// ---- OTEL/TRACING/TRACESTATE/FUNCTION_BLOCKS/TraceStateFactory.TcPOU
(*
	Creates FB_TraceState values: parses a W3C tracestate header, clones a trace state, and
	truncates one to fit a carrier by the W3C rules. Like ValueFactory, every method returns
	TRUE on success, takes pDest by reference and never overwrites a pointer that is not 0.
	No trace state is a 0 pointer, so a method can succeed and leave pDest at 0.
*)
PROGRAM TraceStateFactory
VAR CONSTANT
	MAX_ENTRIES: UDINT := 32;  // W3C: at most 32 list members
	MAX_KEY_LENGTH: UDINT := 256;  // W3C key grammar
	MAX_VALUE_LENGTH: UDINT := 256;  // W3C value grammar
	MAX_HEADER_LENGTH: UDINT := 16447;  // 32 entries of the longest key and value; bounds every scan
	CARRIER_LENGTH: UDINT := 512;  // W3C: propagate at least 512 characters
	LARGE_ENTRY_LENGTH: UDINT := 128;  // W3C: when truncating, remove entries over 128 characters first
END_VAR

(*
	Allocates a trace state from the kept entries of pSource, joined by ','. Succeeds with pDest
	left at 0 when no entry is kept. The arrays are primitive scratch data owned by the caller.
*)
METHOD _build : BOOL
VAR_IN_OUT
	pDest: POINTER TO FB_TraceState;
	starts: ARRAY[0..MAX_ENTRIES - 1] OF UDINT;
	lengths: ARRAY[0..MAX_ENTRIES - 1] OF UDINT;
	keep: ARRAY[0..MAX_ENTRIES - 1] OF BOOL;
END_VAR
VAR_INPUT
	pSource: POINTER TO BYTE;
	count: UDINT;
END_VAR
VAR_OUTPUT
	failureReason: E_TraceStateFailureReason;
END_VAR
VAR
	_i: UDINT;
	_kept: UDINT;
	_length: UDINT;
	_offset: UDINT;
	_pBuffer: POINTER TO BYTE;
	_size: UDINT;
	_pNew: POINTER TO FB_TraceState;
END_VAR
_build := FALSE;
failureReason := E_TraceStateFailureReason.NA;

// size the buffer to the kept entries and the commas between them
WHILE _i < count AND _i < MAX_ENTRIES DO
	IF keep[_i] THEN
		_length := _length + lengths[_i];
		_kept := _kept + 1;
	END_IF
	_i := _i + 1;
END_WHILE
IF _kept = 0 THEN
	// nothing left is no trace state, not an empty one
	_build := TRUE;
	RETURN;
END_IF
_length := _length + _kept - 1;

_size := _length + 1;
_pBuffer := __NEW(BYTE, _size);
IF _pBuffer = 0 THEN
	failureReason := E_TraceStateFailureReason.MEMORY_ALLOCATION_FAILURE;
	RETURN;
END_IF

_i := 0;
WHILE _i < count AND _i < MAX_ENTRIES DO
	IF keep[_i] THEN
		IF _offset > 0 THEN
			_pBuffer[_offset] := 16#2C;  // ','
			_offset := _offset + 1;
		END_IF
		MEMCPY(_pBuffer + _offset, pSource + starts[_i], lengths[_i]);
		_offset := _offset + lengths[_i];
	END_IF
	_i := _i + 1;
END_WHILE
_pBuffer[_offset] := 0;

_pNew := __NEW(FB_TraceState(pString:=_pBuffer, length:=_length, count:=_kept));
IF _pNew = 0 THEN
	__DELETE(_pBuffer);
	_pBuffer := 0;
	failureReason := E_TraceStateFailureReason.MEMORY_ALLOCATION_FAILURE;
	RETURN;
END_IF
pDest := _pNew;
_build := TRUE;
END_METHOD

(* lcalpha / DIGIT / '_' / '-' / '*' / '/' *)
METHOD _isKeyChar : BOOL
VAR_INPUT
	c: BYTE;
END_VAR
_isKeyChar := (c >= 16#61 AND c <= 16#7A)  // a-z
	OR (c >= 16#30 AND c <= 16#39)  // 0-9
	OR c = 16#5F OR c = 16#2D OR c = 16#2A OR c = 16#2F;
END_METHOD

(*
	A key is either simple-key, a lower-case letter followed by up to 255 key characters, or
	multi-tenant-key: tenant-id '@' system-id, where tenant-id is 1-241 key characters starting
	with a lower-case letter or digit, and system-id is 1-14 key characters starting with a
	lower-case letter.
*)
METHOD _isValidKey : BOOL
VAR_INPUT
	pKey: POINTER TO BYTE;
	length: UDINT;
END_VAR
VAR
	_i: UDINT;
	_at: UDINT;
	_hasAt: BOOL;
	_first: BYTE;
END_VAR
_isValidKey := FALSE;
IF length = 0 OR length > MAX_KEY_LENGTH THEN
	RETURN;
END_IF

// bounded by MAX_KEY_LENGTH
WHILE _i < length DO
	IF pKey[_i] = 16#40 THEN  // '@'
		IF _hasAt THEN
			RETURN;
		END_IF
		_hasAt := TRUE;
		_at := _i;
	ELSIF NOT TraceStateFactory._isKeyChar(c:=pKey[_i]) THEN
		RETURN;
	END_IF
	_i := _i + 1;
END_WHILE

_first := pKey[0];
IF NOT _hasAt THEN
	_isValidKey := _first >= 16#61 AND _first <= 16#7A;
ELSIF _at >= 1 AND _at <= 241 AND length - _at - 1 >= 1 AND length - _at - 1 <= 14 THEN
	_isValidKey := ((_first >= 16#61 AND _first <= 16#7A) OR (_first >= 16#30 AND _first <= 16#39))
		AND pKey[_at + 1] >= 16#61 AND pKey[_at + 1] <= 16#7A;
END_IF
END_METHOD

(*
	A value is 1-256 printable ASCII characters other than ',' and '=', and does not end in a
	space.
*)
METHOD _isValidValue : BOOL
VAR_INPUT
	pValue: POINTER TO BYTE;
	length: UDINT;
END_VAR
VAR
	_i: UDINT;
	_c: BYTE;
END_VAR
_isValidValue := FALSE;
IF length = 0 OR length > MAX_VALUE_LENGTH THEN
	RETURN;
END_IF
IF pValue[length - 1] = 16#20 THEN
	RETURN;
END_IF

// bounded by MAX_VALUE_LENGTH
WHILE _i < length DO
	_c := pValue[_i];
	IF _c < 16#20 OR _c > 16#7E OR _c = 16#2C OR _c = 16#3D THEN
		RETURN;
	END_IF
	_i := _i + 1;
END_WHILE
_isValidValue := TRUE;
END_METHOD

(*
	Allocates a copy of pSrc. The caller owns pDest.
*)
METHOD clone : BOOL
VAR_IN_OUT
	pDest: POINTER TO FB_TraceState;
END_VAR
VAR_INPUT
	pSrc: POINTER TO FB_TraceState;
END_VAR
VAR_OUTPUT
	failureReason: E_TraceStateFailureReason;
END_VAR
VAR
	_pBuffer: POINTER TO BYTE;
	_size: UDINT;
	_pNew: POINTER TO FB_TraceState;
END_VAR
clone := FALSE;
failureReason := E_TraceStateFailureReason.NA;

IF pDest <> 0 THEN
	failureReason := E_TraceStateFailureReason.DESTINATION_ALREADY_ASSIGNED;
	RETURN;
END_IF
IF pSrc = 0 OR_ELSE pSrc^.pString = 0 THEN
	failureReason := E_TraceStateFailureReason.SOURCE_POINTER_NULL;
	RETURN;
END_IF

// copy by length, terminator included; the string may be longer than T_MaxString
_size := pSrc^.length + 1;
_pBuffer := __NEW(BYTE, _size);
IF _pBuffer = 0 THEN
	failureReason := E_TraceStateFailureReason.MEMORY_ALLOCATION_FAILURE;
	RETURN;
END_IF
MEMCPY(_pBuffer, pSrc^.pString, pSrc^.length + 1);

_pNew := __NEW(FB_TraceState(pString:=_pBuffer, length:=pSrc^.length, count:=pSrc^.count));
IF _pNew = 0 THEN
	__DELETE(_pBuffer);
	_pBuffer := 0;
	failureReason := E_TraceStateFailureReason.MEMORY_ALLOCATION_FAILURE;
	RETURN;
END_IF
pDest := _pNew;
clone := TRUE;
END_METHOD

(*
	Parses a W3C tracestate header into a new trace state in canonical form. The caller owns
	pDest. An empty header, or one of only empty members, is valid and succeeds with pDest left
	at 0. A header that breaks the grammar, repeats a key or has more than MAX_ENTRIES entries
	fails, and W3C says it must then not be propagated. The header may be longer than
	T_MaxString; it is measured with LEN2.
*)
METHOD parse : BOOL
VAR_IN_OUT
	pDest: POINTER TO FB_TraceState;
END_VAR
VAR_INPUT
	pHeader: POINTER TO STRING;
END_VAR
VAR_OUTPUT
	failureReason: E_TraceStateFailureReason;
END_VAR
VAR
	_pHeader: POINTER TO BYTE;
	_length: UDINT;
	_i: UDINT;
	_j: UDINT;
	_memberStart: UDINT;
	_start: UDINT;
	_end: UDINT;
	_equals: UDINT;
	_keyLength: UDINT;
	_count: UDINT;
	_starts: ARRAY[0..MAX_ENTRIES - 1] OF UDINT;
	_lengths: ARRAY[0..MAX_ENTRIES - 1] OF UDINT;
	_keyLengths: ARRAY[0..MAX_ENTRIES - 1] OF UDINT;
	_keep: ARRAY[0..MAX_ENTRIES - 1] OF BOOL;
END_VAR
parse := FALSE;
failureReason := E_TraceStateFailureReason.NA;

IF pDest <> 0 THEN
	failureReason := E_TraceStateFailureReason.DESTINATION_ALREADY_ASSIGNED;
	RETURN;
END_IF
IF pHeader = 0 THEN
	failureReason := E_TraceStateFailureReason.HEADER_POINTER_NULL;
	RETURN;
END_IF

_pHeader := pHeader;
_length := TO_UDINT(LEN2(pHeader));
IF _length > MAX_HEADER_LENGTH THEN
	failureReason := E_TraceStateFailureReason.HEADER_TOO_LONG;
	RETURN;
END_IF

// validate every member before allocating anything; _i = _length closes the last member
FOR _i := 0 TO _length DO
	IF _i < _length AND_THEN _pHeader[_i] <> 16#2C THEN  // ','
		CONTINUE;
	END_IF
	_start := _memberStart;
	_end := _i;
	_memberStart := _i + 1;

	// strip optional whitespace; an empty member is allowed and dropped
	WHILE _start < _end AND_THEN (_pHeader[_start] = 16#20 OR _pHeader[_start] = 16#09) DO
		_start := _start + 1;
	END_WHILE
	WHILE _end > _start AND_THEN (_pHeader[_end - 1] = 16#20 OR _pHeader[_end - 1] = 16#09) DO
		_end := _end - 1;
	END_WHILE
	IF _start = _end THEN
		CONTINUE;
	END_IF

	IF _count >= MAX_ENTRIES THEN
		failureReason := E_TraceStateFailureReason.TOO_MANY_ENTRIES;
		RETURN;
	END_IF

	_equals := _start;
	WHILE _equals < _end AND_THEN _pHeader[_equals] <> 16#3D DO  // '='
		_equals := _equals + 1;
	END_WHILE
	_keyLength := _equals - _start;
	IF NOT TraceStateFactory._isValidKey(pKey:=_pHeader + _start, length:=_keyLength) THEN
		failureReason := E_TraceStateFailureReason.INVALID_KEY;
		RETURN;
	END_IF
	IF _equals = _end OR_ELSE NOT TraceStateFactory._isValidValue(pValue:=_pHeader + _equals + 1, length:=_end - _equals - 1) THEN
		failureReason := E_TraceStateFailureReason.INVALID_VALUE;
		RETURN;
	END_IF

	_j := 0;
	WHILE _j < _count DO
		IF _keyLengths[_j] = _keyLength AND_THEN MEMCMP(_pHeader + _starts[_j], _pHeader + _start, _keyLength) = 0 THEN
			failureReason := E_TraceStateFailureReason.DUPLICATE_KEY;
			RETURN;
		END_IF
		_j := _j + 1;
	END_WHILE

	_starts[_count] := _start;
	_lengths[_count] := _end - _start;
	_keyLengths[_count] := _keyLength;
	_keep[_count] := TRUE;
	_count := _count + 1;
END_FOR

parse := TraceStateFactory._build(
	pDest:=pDest,
	starts:=_starts,
	lengths:=_lengths,
	keep:=_keep,
	pSource:=_pHeader,
	count:=_count,
	failureReason=>failureReason
);
END_METHOD

(*
	Allocates a copy of pSrc that is at most maxLength characters long, for a carrier of
	limited size, following W3C: entries over LARGE_ENTRY_LENGTH characters are removed first,
	then entries are removed from the right. An entry is removed whole, never cut. Succeeds with
	pDest left at 0 when no entry fits.
*)
METHOD truncate : BOOL
VAR_IN_OUT
	pDest: POINTER TO FB_TraceState;
END_VAR
VAR_INPUT
	pSrc: POINTER TO FB_TraceState;
	maxLength: UDINT;
END_VAR
VAR_OUTPUT
	failureReason: E_TraceStateFailureReason;
END_VAR
VAR
	_pSource: POINTER TO BYTE;
	_i: UDINT;
	_start: UDINT;
	_count: UDINT;
	_kept: UDINT;
	_sum: UDINT;
	_total: UDINT;
	_starts: ARRAY[0..MAX_ENTRIES - 1] OF UDINT;
	_lengths: ARRAY[0..MAX_ENTRIES - 1] OF UDINT;
	_keep: ARRAY[0..MAX_ENTRIES - 1] OF BOOL;
END_VAR
truncate := FALSE;
failureReason := E_TraceStateFailureReason.NA;

IF pDest <> 0 THEN
	failureReason := E_TraceStateFailureReason.DESTINATION_ALREADY_ASSIGNED;
	RETURN;
END_IF
IF pSrc = 0 OR_ELSE pSrc^.pString = 0 THEN
	failureReason := E_TraceStateFailureReason.SOURCE_POINTER_NULL;
	RETURN;
END_IF

IF pSrc^.length <= maxLength THEN
	truncate := TraceStateFactory.clone(pDest:=pDest, pSrc:=pSrc, failureReason=>failureReason);
	RETURN;
END_IF

// split the canonical string: entries joined by ',', no whitespace, at most MAX_ENTRIES
_pSource := pSrc^.pString;
FOR _i := 0 TO pSrc^.length DO
	IF _i = pSrc^.length OR_ELSE _pSource[_i] = 16#2C THEN
		IF _count < MAX_ENTRIES THEN
			_starts[_count] := _start;
			_lengths[_count] := _i - _start;
			_keep[_count] := TRUE;
			_sum := _sum + _i - _start;
			_count := _count + 1;
		END_IF
		_start := _i + 1;
	END_IF
END_FOR
_kept := _count;
_total := pSrc^.length;

// first remove the large entries, from the right
_i := _count;
WHILE _i > 0 AND _total > maxLength DO
	_i := _i - 1;
	IF _lengths[_i] > LARGE_ENTRY_LENGTH THEN
		_keep[_i] := FALSE;
		_sum := _sum - _lengths[_i];
		_kept := _kept - 1;
		_total := SEL(_kept > 0, 0, _sum + _kept - 1);
	END_IF
END_WHILE

// then any entry, from the right
_i := _count;
WHILE _i > 0 AND _total > maxLength DO
	_i := _i - 1;
	IF _keep[_i] THEN
		_keep[_i] := FALSE;
		_sum := _sum - _lengths[_i];
		_kept := _kept - 1;
		_total := SEL(_kept > 0, 0, _sum + _kept - 1);
	END_IF
END_WHILE

truncate := TraceStateFactory._build(
	pDest:=pDest,
	starts:=_starts,
	lengths:=_lengths,
	keep:=_keep,
	pSource:=_pSource,
	count:=_count,
	failureReason=>failureReason
);
END_METHOD

END_PROGRAM

// ---- OTEL/TRACING/SPAN/ContextFactory.TcPOU
PROGRAM ContextFactory

(*
	Allocates a span context holding copies of the given identity. The caller owns pDest.
	The identifiers are not validated; producers are responsible for what they build,
	and a context built from all-zero identifiers is simply not valid.
	pTraceState is borrowed and copied; 0 means no trace state.
*)
METHOD buildContext : BOOL
VAR_IN_OUT
	pDest: POINTER TO FB_SpanContext;
END_VAR
VAR_INPUT
	pTraceId: POINTER TO FB_TraceId;
	pSpanId: POINTER TO FB_SpanId;
	pTraceState: POINTER TO FB_TraceState;
	traceFlags: UDINT;
END_VAR
VAR_OUTPUT
	failureReason: E_ContextFactoryFailureReason;
END_VAR
VAR
	_pTraceState: POINTER TO FB_TraceState;
	_pNew: POINTER TO FB_SpanContext;
END_VAR
buildContext := FALSE;
failureReason := E_ContextFactoryFailureReason.NA;

IF pDest <> 0 THEN
	failureReason := E_ContextFactoryFailureReason.DESTINATION_ALREADY_ASSIGNED;
	RETURN;
END_IF

IF pTraceId = 0 THEN
	failureReason := E_ContextFactoryFailureReason.TRACE_ID_POINTER_NULL;
	RETURN;
END_IF

IF pSpanId = 0 THEN
	failureReason := E_ContextFactoryFailureReason.SPAN_ID_POINTER_NULL;
	RETURN;
END_IF

// clone all owned data before allocating the context itself
IF pTraceState <> 0 THEN
	IF NOT TraceStateFactory.clone(pDest:=_pTraceState, pSrc:=pTraceState) THEN
		failureReason := E_ContextFactoryFailureReason.MEMORY_ALLOCATION_FAILURE;
		RETURN;
	END_IF
END_IF

_pNew := __NEW(FB_SpanContext(
	pTraceId:=pTraceId,
	pSpanId:=pSpanId,
	pTraceState:=_pTraceState,
	traceFlags:=traceFlags
));
IF _pNew = 0 THEN
	failureReason := E_ContextFactoryFailureReason.MEMORY_ALLOCATION_FAILURE;
	IF _pTraceState <> 0 THEN _pTraceState^.delete(pSelf:=_pTraceState); END_IF
	RETURN;
END_IF
_pTraceState := 0;  // moved into FB_SpanContext
pDest := _pNew;
buildContext := failureReason = E_ContextFactoryFailureReason.NA;
END_METHOD

(*
	Allocates a snapshot of a span's identity. The caller owns pDest, which must be 0; the span
	is borrowed and unchanged. The span is the producer, and its identifiers come from the id
	generator, which only hands out valid ones, so they are not checked again here. A span that
	has not been built has no identifiers and is refused with TRACE_ID_POINTER_NULL.
	The context is always local: a span's own flags describe its parent's remoteness, so only
	the W3C trace flags are kept, and remoteness is marked as known and not remote.
*)
METHOD fromSpan : BOOL
VAR_IN_OUT
	pDest: POINTER TO FB_SpanContext;
END_VAR
VAR_INPUT
	pSpan: POINTER TO FB_Span;
END_VAR
VAR_OUTPUT
	failureReason: E_ContextFactoryFailureReason;
END_VAR
VAR
	_traceFlags: UDINT;
END_VAR
fromSpan := FALSE;
failureReason := E_ContextFactoryFailureReason.NA;

IF pSpan = 0 THEN
	failureReason := E_ContextFactoryFailureReason.SPAN_POINTER_NULL;
	RETURN;
END_IF

_traceFlags := (pSpan^.flags AND TO_UDINT(E_SpanFlags.SPAN_FLAGS_TRACE_FLAGS_MASK))
	OR TO_UDINT(E_SpanFlags.SPAN_FLAGS_CONTEXT_HAS_IS_REMOTE_MASK);

fromSpan := ContextFactory.buildContext(
	pDest:=pDest,
	pTraceId:=pSpan^.traceId,
	pSpanId:=pSpan^.spanId,
	pTraceState:=pSpan^.traceState,
	traceFlags:=_traceFlags,
	failureReason=>failureReason
);
END_METHOD

END_PROGRAM

// ---- OTEL/COMMON/FUNCTION_BLOCKS/FB_Resource.TcPOU
{attribute 'enable_dynamic_creation'}
FUNCTION_BLOCK FB_Resource
VAR_OUTPUT
	id: UDINT;	// process-local identity, assigned automatically and never exported. Snapshots share the id of their source.
	droppedAttributesCount: UDINT;
	schemaUrl: T_MaxString;
END_VAR
VAR_OUTPUT
	attributes: FB_Attributes(maxCount := TcOtlp_GVL.DEFAULT_MAX_ATTRIBUTE_COUNT);
END_VAR

METHOD copyFrom : BOOL
VAR_IN_OUT
	src: FB_Resource;
END_VAR
VAR_OUTPUT
	failureResult: E_AttributesFailureReason;
END_VAR
failureResult := E_AttributesFailureReason.NA;
THIS^.id := src.id;
THIS^.schemaUrl := src.schemaUrl;
THIS^.droppedAttributesCount := src.droppedAttributesCount;
THIS^.attributes.free();
copyFrom := THIS^.attributes.copyFrom(src:=src.attributes, failureReason=>failureResult);
END_METHOD

METHOD FB_Exit : BOOL
VAR_INPUT
	bInCopyCode: BOOL;
END_VAR
THIS^.free();
END_METHOD

//FB_Init is always available implicitly and it is used primarily for initialization.
//The return value is not evaluated. For a specific influence, you can also declare the
//methods explicitly and provide additional code there with the standard initialization
//code. You can evaluate the return value.
METHOD FB_Init: BOOL
VAR_INPUT
    bInitRetains: BOOL; // TRUE: the retain variables are initialized (reset warm / reset cold)
    bInCopyCode: BOOL;  // TRUE: the instance will be copied to the copy code afterward (online change) 
	schemaUrl: T_MaxString;
END_VAR
THIS^.schemaUrl := schemaUrl;

// claim a process-local identity; keep the existing one during an online change copy
IF NOT bInCopyCode THEN
	THIS^.id := TcOtlp_GVL.NEXT_ID;
END_IF
END_METHOD

METHOD free
THIS^.attributes.free();
END_METHOD

END_FUNCTION_BLOCK

// ---- OTEL/COMMON/FUNCTION_BLOCKS/FB_InstrumentationScope.TcPOU
FUNCTION_BLOCK FB_InstrumentationScope
VAR_OUTPUT
	name: T_MaxString;
	version: T_MaxString;
	droppedAttributesCount: UDINT;
	schemaUrl: T_MaxString;
END_VAR
VAR_OUTPUT
	attributes: FB_Attributes(maxCount := TcOtlp_GVL.DEFAULT_MAX_ATTRIBUTE_COUNT);
END_VAR

METHOD copyFrom : BOOL
VAR_IN_OUT
	src: FB_InstrumentationScope;
END_VAR
VAR_OUTPUT
	failureResult: E_AttributesFailureReason;
END_VAR
failureResult := E_AttributesFailureReason.NA;
THIS^.name := src.name;
THIS^.version := src.version;
THIS^.droppedAttributesCount := src.droppedAttributesCount;
THIS^.schemaUrl := src.schemaUrl;
THIS^.attributes.free();
copyFrom := THIS^.attributes.copyFrom(src:=src.attributes, failureReason=>failureResult);
END_METHOD

//FB_Exit must be implemented explicitly. If there is an implementation, then the
//method is called before the controller removes the code of the function block instance
//(implicit call). The return value is not evaluated.
METHOD FB_Exit: BOOL
VAR_INPUT
    bInCopyCode: BOOL;  // TRUE: the exit method is called in order to leave the instance which will be copied afterwards (online change).  
END_VAR
THIS^.free();
END_METHOD

METHOD FB_Init: BOOL
VAR_INPUT
	bInitRetains: BOOL;
	bInCopyCode: BOOL;
	name: T_MaxString;
	version: T_MaxString;
	schemaUrl: T_MaxString;
END_VAR
THIS^.name := name;
THIS^.version := version;
THIS^.schemaUrl := schemaUrl;
END_METHOD

METHOD free
VAR_INPUT
END_VAR
THIS^.attributes.free();
END_METHOD

END_FUNCTION_BLOCK

// ---- OTEL/LOGGING/EXPORTING/FUNCTION_BLOCKS/FB_LogRecordExporter_Base.TcPOU
FUNCTION_BLOCK ABSTRACT FB_LogRecordExporter_Base
VAR
	_records: FB_LogRecordQueue(maxCount:=0);
	_exportActive: BOOL;
	_callFailureReason: E_LogRecordExporterFailureReason;
END_VAR

METHOD export: BOOL
VAR_IN_OUT
	logRecords: FB_LogRecordQueue;  // accepted records are transferred out of this queue
END_VAR
VAR_INPUT
	count: UDINT;
END_VAR
VAR_OUTPUT
	failureReason: E_LogRecordExporterFailureReason;
END_VAR
VAR
	_queueFailureReason: E_LogRecordQueueFailureReason;
END_VAR
export := FALSE;
failureReason := E_LogRecordExporterFailureReason.NA;

IF THIS^.isBusy() THEN
	failureReason := E_LogRecordExporterFailureReason.ACTIVE_EXPORT_IN_PROGRESS;
	RETURN;
END_IF

// Release a completed batch retained by an exporter before accepting the next one.
THIS^.free();
IF NOT logRecords.transferTo(
	destination:=THIS^._records,
	count:=count,
	failureReason=>_queueFailureReason
) THEN
	failureReason := E_LogRecordExporterFailureReason.QUEUE_TRANSFER_FAILURE;
	RETURN;
END_IF

THIS^._exportActive := THIS^._records.count > 0;
export := failureReason = E_LogRecordExporterFailureReason.NA;
END_METHOD

METHOD FB_Exit: BOOL
VAR_INPUT
	bInCopyCode: BOOL;
END_VAR
IF NOT bInCopyCode THEN
	THIS^.free();
END_IF
END_METHOD

METHOD free
THIS^._records.free();
THIS^._exportActive := FALSE;
END_METHOD

METHOD ABSTRACT isBusy : BOOL
END_METHOD

METHOD ABSTRACT tick : BOOL
VAR_OUTPUT
	failureReason: E_LogRecordExporterFailureReason;
END_VAR
END_METHOD

END_FUNCTION_BLOCK

// ---- OTEL/LOGGING/LOG_RECORD/FUNCTION_BLOCKS/FB_LogRecordQueue.TcPOU
(*
	FIFO queue that owns every FB_LogRecord pointer it contains. push drops the
	oldest owned records when the bound is reached. The bound is maxCount, but
	never more than TcOtlp_GVL.MAX_LOOP_COUNT: a maxCount of zero, or one above
	that limit, is held to MAX_LOOP_COUNT so that free always reaches the end.
	pop transfers ownership back to the caller. transferTo moves allocated
	nodes between queue owners without copying records.
*)
FUNCTION_BLOCK FB_LogRecordQueue
VAR
	_head: POINTER TO ST_LinkedListNode;
	_tail: POINTER TO ST_LinkedListNode;
	_cursor: POINTER TO ST_LinkedListNode;
END_VAR
VAR_OUTPUT
	count: UDINT;
	maxCount: UDINT;
	droppedCount: UDINT;
END_VAR

(* The enforced bound: maxCount, held to MAX_LOOP_COUNT when it is zero or larger. *)
METHOD _capacity : UDINT
IF THIS^.maxCount = 0 OR THIS^.maxCount > TcOtlp_GVL.MAX_LOOP_COUNT THEN
	_capacity := TcOtlp_GVL.MAX_LOOP_COUNT;
ELSE
	_capacity := THIS^.maxCount;
END_IF
END_METHOD

METHOD FB_Exit : BOOL
VAR_INPUT
	bInCopyCode: BOOL;
END_VAR
IF NOT bInCopyCode THEN
	THIS^.free();
END_IF
END_METHOD

METHOD FB_Init : BOOL
VAR_INPUT
	bInitRetains: BOOL;
	bInCopyCode: BOOL;
	maxCount: UDINT := 0;
END_VAR
THIS^.maxCount := maxCount;
END_METHOD

(*
	Releases every owned record. push holds count to MAX_LOOP_COUNT, so the loop
	always reaches the end. If it ever stops early, the unreleased nodes stay in
	the queue and free returns FALSE, so a later call can finish the job.
*)
METHOD free : BOOL
VAR
	_idx: UDINT;
	_node: POINTER TO ST_LinkedListNode;
	_record: POINTER TO FB_LogRecord;
END_VAR
FOR _idx := 0 TO TcOtlp_GVL.MAX_LOOP_COUNT DO
	IF THIS^._head = 0 THEN
		EXIT;
	END_IF

	_node := THIS^._head;
	THIS^._head := _node^.nxt;
	IF _node^.val <> 0 THEN
		_record := _node^.val;
		_node^.val := 0;
		_record^.delete(pSelf:=_record);
	END_IF
	__DELETE(_node);
	IF THIS^.count > 0 THEN
		THIS^.count := THIS^.count - 1;
	END_IF
END_FOR

THIS^._cursor := THIS^._head;
IF THIS^._head = 0 THEN
	THIS^._tail := 0;
	THIS^.count := 0;
END_IF
free := THIS^._head = 0;
END_METHOD

METHOD next : POINTER TO FB_LogRecord
next := 0;

IF THIS^._cursor <> 0 THEN
	next := THIS^._cursor^.val;
	THIS^._cursor := THIS^._cursor^.nxt;
END_IF
END_METHOD

METHOD pop : BOOL
VAR_IN_OUT
	pValue: POINTER TO FB_LogRecord;
END_VAR
VAR_OUTPUT
	failureReason: E_LogRecordQueueFailureReason;
END_VAR
VAR
	_node: POINTER TO ST_LinkedListNode;
END_VAR
pop := FALSE;
failureReason := E_LogRecordQueueFailureReason.NA;

IF pValue <> 0 THEN
	failureReason := E_LogRecordQueueFailureReason.DESTINATION_ALREADY_ASSIGNED;
	RETURN;
END_IF
IF THIS^._head = 0 THEN
	failureReason := E_LogRecordQueueFailureReason.QUEUE_EMPTY;
	RETURN;
END_IF

_node := THIS^._head;
THIS^._head := _node^.nxt;
IF THIS^._cursor = _node THEN
	THIS^._cursor := THIS^._head;
END_IF
IF THIS^._head = 0 THEN
	THIS^._tail := 0;
END_IF

pValue := _node^.val;
_node^.val := 0;
_node^.nxt := 0;
__DELETE(_node);
_node := 0;
THIS^.count := THIS^.count - 1;
pop := failureReason = E_LogRecordQueueFailureReason.NA;
END_METHOD

METHOD push : BOOL
VAR_IN_OUT
	pValue: POINTER TO FB_LogRecord;
END_VAR
VAR_OUTPUT
	failureReason: E_LogRecordQueueFailureReason;
END_VAR
VAR
	_node: POINTER TO ST_LinkedListNode;
	_droppedRecord: POINTER TO FB_LogRecord;
	_popFailureReason: E_LogRecordQueueFailureReason;
	_idx: UDINT;
	_bound: UDINT;
END_VAR
push := FALSE;
failureReason := E_LogRecordQueueFailureReason.NA;

IF pValue = 0 THEN
	failureReason := E_LogRecordQueueFailureReason.RECORD_POINTER_NULL;
	RETURN;
END_IF

// Allocate before evicting so an allocation failure leaves the queue unchanged.
_node := __NEW(ST_LinkedListNode);
IF _node = 0 THEN
	failureReason := E_LogRecordQueueFailureReason.MEMORY_ALLOCATION_FAILURE;
	RETURN;
END_IF

// maxCount is writable, so also restore the bound after a runtime reduction.
_bound := THIS^._capacity();
FOR _idx := 0 TO TcOtlp_GVL.MAX_LOOP_COUNT DO
	IF THIS^.count < _bound THEN
		EXIT;
	END_IF
	IF NOT THIS^.pop(pValue:=_droppedRecord, failureReason=>_popFailureReason) THEN
		__DELETE(_node);
		_node := 0;
		failureReason := _popFailureReason;
		RETURN;
	END_IF
	_droppedRecord^.delete(pSelf:=_droppedRecord);
	THIS^.droppedCount := THIS^.droppedCount + 1;
END_FOR
IF THIS^.count >= _bound THEN
	__DELETE(_node);
	_node := 0;
	failureReason := E_LogRecordQueueFailureReason.MAX_SIZE_ENFORCEMENT_FAILURE;
	RETURN;
END_IF

_node^.val := pValue;
_node^.nxt := 0;
IF THIS^._tail = 0 THEN
	THIS^._head := _node;
	THIS^._cursor := _node;
ELSE
	THIS^._tail^.nxt := _node;
END_IF
THIS^._tail := _node;
THIS^.count := THIS^.count + 1;
pValue := 0;
push := failureReason = E_LogRecordQueueFailureReason.NA;
END_METHOD

METHOD reset
THIS^._cursor := THIS^._head;
END_METHOD

(* Moves the head node to the tail without changing record ownership. *)
METHOD rotate : BOOL
VAR_OUTPUT
	failureReason: E_LogRecordQueueFailureReason;
END_VAR
VAR
	_node: POINTER TO ST_LinkedListNode;
END_VAR
rotate := FALSE;
failureReason := E_LogRecordQueueFailureReason.NA;

IF THIS^._head = 0 THEN
	failureReason := E_LogRecordQueueFailureReason.QUEUE_EMPTY;
	RETURN;
END_IF

IF THIS^._head <> THIS^._tail THEN
	_node := THIS^._head;
	THIS^._head := _node^.nxt;
	_node^.nxt := 0;
	THIS^._tail^.nxt := _node;
	THIS^._tail := _node;
END_IF

THIS^._cursor := THIS^._head;
rotate := failureReason = E_LogRecordQueueFailureReason.NA;
END_METHOD

(*
	Transfers the allocated nodes and owned records without copying them.
	The destination must be a different, empty queue. It receives up to count
	of the oldest records, also respecting the destination's bound.
*)
METHOD transferTo : BOOL
VAR_IN_OUT
	destination: FB_LogRecordQueue;
END_VAR
VAR_INPUT
	count: UDINT;
END_VAR
VAR_OUTPUT
	failureReason: E_LogRecordQueueFailureReason;
END_VAR
VAR
	_transferCount: UDINT;
	_idx: UDINT;
END_VAR
transferTo := FALSE;
failureReason := E_LogRecordQueueFailureReason.NA;

IF ADR(destination) = THIS THEN
	failureReason := E_LogRecordQueueFailureReason.SELF_TRANSFER_NOT_ALLOWED;
	RETURN;
END_IF
IF destination.count <> 0 OR_ELSE destination._head <> 0 OR_ELSE destination._tail <> 0 THEN
	failureReason := E_LogRecordQueueFailureReason.DESTINATION_NOT_EMPTY;
	RETURN;
END_IF

_transferCount := count;
IF _transferCount > THIS^.count THEN
	_transferCount := THIS^.count;
END_IF
IF _transferCount > destination._capacity() THEN
	_transferCount := destination._capacity();
END_IF
IF _transferCount = 0 THEN
	transferTo := failureReason = E_LogRecordQueueFailureReason.NA;
	RETURN;
END_IF

destination._head := THIS^._head;
destination._tail := destination._head;
FOR _idx := 1 TO _transferCount - 1 DO
	destination._tail := destination._tail^.nxt;
END_FOR

THIS^._head := destination._tail^.nxt;
destination._tail^.nxt := 0;
destination._cursor := destination._head;
destination.count := _transferCount;

THIS^.count := THIS^.count - _transferCount;
THIS^._cursor := THIS^._head;
IF THIS^._head = 0 THEN
	THIS^._tail := 0;
END_IF
transferTo := failureReason = E_LogRecordQueueFailureReason.NA;
END_METHOD

END_FUNCTION_BLOCK

// ---- OTEL/LOGGING/LOG_RECORD/FUNCTION_BLOCKS/FB_LogRecord.TcPOU
{attribute 'enable_dynamic_creation'}
FUNCTION_BLOCK FB_LogRecord
VAR_INPUT
	// required values
	severityNumber: E_SeverityNumber;
	timestamp: 		ULINT;
	
	// optional values
	eventName: 	POINTER TO FB_String; 
	traceId: 	POINTER TO FB_TraceId;
	spanId: 	POINTER TO FB_SpanId;
	flags: UDINT;  // OTLP fixed32: bits 0-7 are the W3C trace flags of the record's span (bit 0 is sampled), bits 8-31 are reserved
	body: 		POINTER TO FB_AnyValue;
	droppedAttributesCount: UDINT;
END_VAR
VAR_OUTPUT
	resource: FB_Resource('');
	scope: FB_InstrumentationScope('', '', '');
	attributes: FB_Attributes(maxCount := TcOtlp_GVL.DEFAULT_MAX_ATTRIBUTE_COUNT);
END_VAR

METHOD cloneTo : BOOL
VAR_IN_OUT
	pDest: POINTER TO FB_LogRecord;
END_VAR
VAR_OUTPUT
	failureReason: E_LogRecordCloneFailureReason;
END_VAR
VAR
	_pClone: POINTER TO FB_LogRecord;
	_factoryFailureReason: E_ValueFactoryFailureReason;
	_attributesFailureReason: E_AttributesFailureReason;
END_VAR
cloneTo := FALSE;
failureReason := E_LogRecordCloneFailureReason.NA;

IF pDest <> 0 THEN
	failureReason := E_LogRecordCloneFailureReason.DESTINATION_ALREADY_ASSIGNED;
	RETURN;
END_IF

_pClone := __NEW(FB_LogRecord(
	severityNumber:=THIS^.severityNumber,
	timestamp:=THIS^.timestamp
));
IF _pClone = 0 THEN
	failureReason := E_LogRecordCloneFailureReason.MEMORY_ALLOCATION_FAILURE;
	RETURN;
END_IF

_pClone^.droppedAttributesCount := THIS^.droppedAttributesCount;
_pClone^.flags := THIS^.flags;

IF THIS^.eventName <> 0 THEN
	IF NOT ValueFactory.cloneString(
		pDest:=_pClone^.eventName,
		pSrc:=THIS^.eventName,
		failureReason=>_factoryFailureReason
	) THEN
		IF _factoryFailureReason = E_ValueFactoryFailureReason.MEMORY_ALLOCATION_FAILURE THEN
			failureReason := E_LogRecordCloneFailureReason.MEMORY_ALLOCATION_FAILURE;
		ELSE
			failureReason := E_LogRecordCloneFailureReason.EVENT_NAME_INVALID;
		END_IF
		_pClone^.delete(pSelf:=_pClone);
		RETURN;
	END_IF
END_IF

IF THIS^.traceId <> 0 THEN
	IF NOT ValueFactory.createTraceId(
		pDest:=_pClone^.traceId,
		pBytes:=ADR(THIS^.traceId^.bytes),
		nSize:=SIZEOF(THIS^.traceId^.bytes),
		failureReason=>_factoryFailureReason
	) THEN
		IF _factoryFailureReason = E_ValueFactoryFailureReason.MEMORY_ALLOCATION_FAILURE THEN
			failureReason := E_LogRecordCloneFailureReason.MEMORY_ALLOCATION_FAILURE;
		ELSE
			failureReason := E_LogRecordCloneFailureReason.TRACE_ID_INVALID;
		END_IF
		_pClone^.delete(pSelf:=_pClone);
		RETURN;
	END_IF
END_IF

IF THIS^.spanId <> 0 THEN
	IF NOT ValueFactory.createSpanId(
		pDest:=_pClone^.spanId,
		pBytes:=ADR(THIS^.spanId^.bytes),
		nSize:=SIZEOF(THIS^.spanId^.bytes),
		failureReason=>_factoryFailureReason
	) THEN
		IF _factoryFailureReason = E_ValueFactoryFailureReason.MEMORY_ALLOCATION_FAILURE THEN
			failureReason := E_LogRecordCloneFailureReason.MEMORY_ALLOCATION_FAILURE;
		ELSE
			failureReason := E_LogRecordCloneFailureReason.SPAN_ID_INVALID;
		END_IF
		_pClone^.delete(pSelf:=_pClone);
		RETURN;
	END_IF
END_IF

IF THIS^.body <> 0 THEN
	IF NOT ValueFactory.cloneAnyValue(
		pDest:=_pClone^.body,
		pSrc:=THIS^.body,
		failureReason=>_factoryFailureReason
	) THEN
		CASE _factoryFailureReason OF
			E_ValueFactoryFailureReason.MEMORY_ALLOCATION_FAILURE:
				failureReason := E_LogRecordCloneFailureReason.MEMORY_ALLOCATION_FAILURE;
			E_ValueFactoryFailureReason.UNSUPPORTED_VALUE_TYPE:
				failureReason := E_LogRecordCloneFailureReason.BODY_VALUE_TYPE_UNSUPPORTED;
		ELSE
			failureReason := E_LogRecordCloneFailureReason.BODY_VALUE_INVALID;
		END_CASE
		_pClone^.delete(pSelf:=_pClone);
		RETURN;
	END_IF
END_IF

IF NOT _pClone^.resource.copyFrom(src:=THIS^.resource, failureResult=>_attributesFailureReason) THEN
	IF _attributesFailureReason = E_AttributesFailureReason.MEMORY_ALLOCATION_FAILURE THEN
		failureReason := E_LogRecordCloneFailureReason.MEMORY_ALLOCATION_FAILURE;
	ELSE
		failureReason := E_LogRecordCloneFailureReason.RESOURCE_COPY_FAILURE;
	END_IF
	_pClone^.delete(pSelf:=_pClone);
	RETURN;
END_IF

IF NOT _pClone^.scope.copyFrom(src:=THIS^.scope, failureResult=>_attributesFailureReason) THEN
	IF _attributesFailureReason = E_AttributesFailureReason.MEMORY_ALLOCATION_FAILURE THEN
		failureReason := E_LogRecordCloneFailureReason.MEMORY_ALLOCATION_FAILURE;
	ELSE
		failureReason := E_LogRecordCloneFailureReason.SCOPE_COPY_FAILURE;
	END_IF
	_pClone^.delete(pSelf:=_pClone);
	RETURN;
END_IF

IF NOT _pClone^.attributes.copyFrom(
	src:=THIS^.attributes,
	failureReason=>_attributesFailureReason
	) THEN
	IF _attributesFailureReason = E_AttributesFailureReason.MEMORY_ALLOCATION_FAILURE THEN
		failureReason := E_LogRecordCloneFailureReason.MEMORY_ALLOCATION_FAILURE;
	ELSE
		failureReason := E_LogRecordCloneFailureReason.ATTRIBUTE_COPY_FAILURE;
	END_IF
	_pClone^.delete(pSelf:=_pClone);
	RETURN;
END_IF

pDest := _pClone;
_pClone := 0;
cloneTo := failureReason = E_LogRecordCloneFailureReason.NA;
END_METHOD

(*
	Releases this record and clears the caller's pointer to it: call it as p^.delete(pSelf:=p).
	pSelf is cleared before the record is freed, so the caller never keeps a dangling pointer.
	A pointer to any other object is refused and left untouched, and nothing is released.
*)
METHOD delete : BOOL
VAR_IN_OUT
	pSelf: POINTER TO FB_LogRecord;
END_VAR
VAR
	_pThis: POINTER TO FB_LogRecord;
END_VAR
_pThis := THIS;
IF pSelf <> _pThis THEN
	RETURN;
END_IF

pSelf := 0;
__DELETE(_pThis);
delete := TRUE;
END_METHOD

//FB_Exit must be implemented explicitly. If there is an implementation, then the
//method is called before the controller removes the code of the function block instance
//(implicit call). The return value is not evaluated.
METHOD FB_Exit: BOOL
VAR_INPUT
    bInCopyCode: BOOL;  // TRUE: the exit method is called in order to leave the instance which will be copied afterwards (online change).
END_VAR
IF NOT bInCopyCode THEN
	THIS^.free();
END_IF
END_METHOD

//FB_Init is always available implicitly and it is used primarily for initialization.
//The return value is not evaluated. For a specific influence, you can also declare the
//methods explicitly and provide additional code there with the standard initialization
//code. You can evaluate the return value.
METHOD FB_Init: BOOL
VAR_INPUT
    bInitRetains: BOOL; // TRUE: the retain variables are initialized (reset warm / reset cold)
    bInCopyCode: BOOL;  // TRUE: the instance will be copied to the copy code afterward (online change)
	// required values
	severityNumber: E_SeverityNumber;
	timestamp: 		ULINT;
END_VAR
// required values
THIS^.severityNumber := severityNumber;
THIS^.timestamp := timestamp;
END_METHOD

METHOD free
IF THIS^.eventName <> 0 THEN THIS^.eventName^.delete(pSelf:=THIS^.eventName); END_IF
IF THIS^.traceId <> 0 THEN THIS^.traceId^.delete(pSelf:=THIS^.traceId); END_IF
IF THIS^.spanId <> 0 THEN THIS^.spanId^.delete(pSelf:=THIS^.spanId); END_IF
IF THIS^.body <> 0 THEN THIS^.body^.delete(pSelf:=THIS^.body); END_IF
THIS^.attributes.free();
THIS^.scope.free();
THIS^.resource.free();
END_METHOD

PROPERTY severityText : STRING(30)
GET
severityText := TO_STRING(THIS^.severityNumber);
END_GET
END_PROPERTY

END_FUNCTION_BLOCK

// ---- OTEL/LOGGING/EXPORTING/FUNCTION_BLOCKS/FB_LogRecordExporter_Console.TcPOU
FUNCTION_BLOCK FB_LogRecordExporter_Console EXTENDS FB_LogRecordExporter_Base
VAR_INPUT
END_VAR
VAR_OUTPUT
END_VAR
VAR
END_VAR

THIS^.tick(failureReason=>THIS^._callFailureReason);

METHOD export : BOOL
VAR_IN_OUT
	logRecords: FB_LogRecordQueue;
END_VAR
VAR_INPUT
	count: UDINT;
END_VAR
VAR_OUTPUT
	failureReason: E_LogRecordExporterFailureReason;
END_VAR
export := SUPER^.export(
	logRecords:=logRecords,
	count:=count,
	failureReason=>failureReason
);
IF NOT export THEN
	RETURN;
END_IF

THIS^.writeToConsole(THIS^._records);
THIS^.free();
END_METHOD

METHOD isBusy : BOOL
isBusy := FALSE;
END_METHOD

METHOD tick : BOOL
VAR_OUTPUT
	failureReason: E_LogRecordExporterFailureReason;
END_VAR
failureReason := E_LogRecordExporterFailureReason.NA;
tick := TRUE;
END_METHOD

METHOD writeToConsole
VAR_IN_OUT
	logRecords: FB_LogRecordQueue;
END_VAR
VAR
	idx: DINT;
	logRecord: POINTER TO FB_LogRecord;
	body: POINTER TO FB_String;
END_VAR
logRecords.reset();
FOR idx := 0 TO TcOtlp_GVL.MAX_LOOP_COUNT DO
	logRecord := logRecords.next();
	IF logRecord = 0 THEN
		RETURN;
	END_IF
	IF logRecord^.body <> 0 AND_THEN logRecord^.body^.eType = E_ValueType.E_String THEN
		body := logRecord^.body;
		ADSLOGSTR(
			ADSLOG_MSGTYPE_ERROR,
			body^.pString^,
			''
		);
	END_IF
END_FOR
END_METHOD

END_FUNCTION_BLOCK

// ---- OTEL/LOGGING/EXPORTING/FUNCTION_BLOCKS/FB_LogRecordExporter_File.TcPOU
FUNCTION_BLOCK FB_LogRecordExporter_File EXTENDS FB_LogRecordExporter_Base
VAR_INPUT
	// maxFileSize: 	UDINT;  // size at which to auto rotate the file
	// maxFiles: 		UDINT;  // max number of files to keep in the rotation
END_VAR

VAR_OUTPUT
	currentState: E_FileExporterState;
END_VAR

VAR
	_execute: BOOL;
	_filepath: T_MaxString;
	_hFile: UINT;
	_len: UDINT;
	_execRTrig: R_TRIG;
	_pString: POINTER TO STRING;
	_jsonVal: SJsonValue;
	_resourceLogsArray: SJsonValue;
	_fileOpener: FB_FileOpen;
	_fileWriter: FB_FileWrite;
	_fileCloser: FB_FileClose;
	_computedState: E_FileExporterState;
	_failureReason: E_LogRecordExporterFailureReason;
	_serializationFailureReason: E_ProtoJsonSerializerFailureReason;
	_serializer: FB_LogRecordProtoJsonSerializer;
END_VAR

THIS^.tick(failureReason=>THIS^._callFailureReason);

METHOD export: BOOL
VAR_IN_OUT
	logRecords: FB_LogRecordQueue;
END_VAR
VAR_INPUT
	count: UDINT;
END_VAR
VAR_OUTPUT
	failureReason: E_LogRecordExporterFailureReason;
END_VAR
// Prepare a completed exporter to accept the next batch immediately.
IF THIS^.currentState = E_FileExporterState.done OR THIS^.currentState = E_FileExporterState.error THEN
	THIS^.currentState := E_FileExporterState.idle;
	THIS^._computedState := E_FileExporterState.idle;
END_IF
export := SUPER^.export(
	logRecords:=logRecords,
	count:=count,
	failureReason=>failureReason
);
IF export THEN
	THIS^._failureReason := E_LogRecordExporterFailureReason.NA;
	THIS^._serializationFailureReason := E_ProtoJsonSerializerFailureReason.NA;
END_IF
END_METHOD

(*
	Releases a payload buffer that is still in flight. The FB_FileWrite reading it is
	destroyed with this instance, so nothing uses the buffer afterwards. TwinCAT then
	runs FB_LogRecordExporter_Base.FB_Exit, which releases the queued records.
*)
METHOD FB_Exit : BOOL
VAR_INPUT
	bInCopyCode: BOOL;  // TRUE: the instance is being copied during an online change
END_VAR
// during an online change the copy keeps the buffer, so it must not be released here
IF NOT bInCopyCode AND _pString <> 0 THEN
	__DELETE(_pString);
	_pString := 0;
END_IF
END_METHOD

//FB_Init is always available implicitly and it is used primarily for initialization.
//The return value is not evaluated. For a specific influence, you can also declare the
//methods explicitly and provide additional code there with the standard initialization
//code. You can evaluate the return value.
METHOD FB_Init: BOOL
VAR_INPUT
    bInitRetains: BOOL; // TRUE: the retain variables are initialized (reset warm / reset cold)
    bInCopyCode: BOOL;  // TRUE: the instance will be copied to the copy code afterward (online change)
	filepath: T_MaxString;  // path to the root file
END_VAR
THIS^._filepath := filepath;
END_METHOD

METHOD isBusy : BOOL
isBusy := THIS^._exportActive;
END_METHOD

METHOD tick : BOOL
VAR_OUTPUT
	failureReason: E_LogRecordExporterFailureReason;
END_VAR
tick := TRUE;
failureReason := E_LogRecordExporterFailureReason.NA;

_execute := THIS^._exportActive;
_execRTrig(CLK := _execute AND_THEN THIS^._records.count > 0);

CASE currentState OF
	E_FileExporterState.idle:
		IF _execRTrig.Q THEN
			_failureReason := E_LogRecordExporterFailureReason.NA;
			_serializationFailureReason := E_ProtoJsonSerializerFailureReason.NA;
			_computedState := E_FileExporterState.serializing;
		END_IF

	E_FileExporterState.serializing:
		IF NOT _serializer.serializeLogsData(
			logRecords:=THIS^._records,
			failureReason=>_serializationFailureReason
		) THEN
			_failureReason := E_LogRecordExporterFailureReason.SERIALIZATION_FAILURE;
			_computedState := E_FileExporterState.error;
		ELSE
			_jsonVal := _serializer.jsonValue;
			IF _jsonVal = 0 OR_ELSE NOT _serializer.parser.IsObject(_jsonVal) THEN
				_failureReason := E_LogRecordExporterFailureReason.SERIALIZATION_FAILURE;
				_computedState := E_FileExporterState.error;
			ELSE
				_resourceLogsArray := _serializer.parser.FindMember(_jsonVal, 'resourceLogs');
				IF _resourceLogsArray = 0 OR_ELSE NOT _serializer.parser.IsArray(_resourceLogsArray) THEN
					_failureReason := E_LogRecordExporterFailureReason.SERIALIZATION_FAILURE;
					_computedState := E_FileExporterState.error;
				ELSE
					_computedState := E_FileExporterState.opening;
				END_IF
			END_IF
		END_IF

	E_FileExporterState.opening:
		IF _fileOpener.bError THEN
			_failureReason := E_LogRecordExporterFailureReason.FILE_OPEN_FAILURE;
			_computedState := E_FileExporterState.error;
		ELSIF NOT _fileOpener.bBusy THEN
			_hFile := _fileOpener.hFile;
			_computedState := E_FileExporterState.buffering;
		END_IF

	E_FileExporterState.buffering:
		// Write one complete LogsData object per JSONL line.
		_len := _serializer.parser.GetJsonLength(_jsonVal);  // includes the null terminating character
		IF _len = 0 THEN
			_failureReason := E_LogRecordExporterFailureReason.SERIALIZATION_FAILURE;
			_computedState := E_FileExporterState.closing;
		ELSE
			_pString := __NEW(BYTE, (_len + 1));  // + 1 for the new line
			IF _pString = 0 THEN
				_failureReason := E_LogRecordExporterFailureReason.BUFFER_ALLOCATION_FAILURE;
				_computedState := E_FileExporterState.closing;
			ELSE
				_serializer.parser.CopyJson(_jsonVal, _pString^, _len);
				CONCAT2(_pString, ADR('$N'), _pString, _len + 1);
				_computedState := E_FileExporterState.writing;
			END_IF
		END_IF

	E_FileExporterState.writing:
		IF _fileWriter.bError THEN
			IF _pString <> 0 THEN __DELETE(_pString); _pString := 0; END_IF
			_failureReason := E_LogRecordExporterFailureReason.FILE_WRITE_FAILURE;
			_computedState := E_FileExporterState.closing;
		ELSIF NOT _fileWriter.bBusy THEN
			IF _pString <> 0 THEN __DELETE(_pString); _pString := 0; END_IF
			_computedState := E_FileExporterState.closing;
		END_IF

	E_FileExporterState.closing:
		IF _fileCloser.bError THEN
			IF _failureReason = E_LogRecordExporterFailureReason.NA THEN
				_failureReason := E_LogRecordExporterFailureReason.FILE_CLOSE_FAILURE;
			END_IF
			_computedState := E_FileExporterState.error;
		ELSIF NOT _fileCloser.bBusy THEN
			IF _failureReason = E_LogRecordExporterFailureReason.NA THEN
				_computedState := E_FileExporterState.done;
			ELSE
				_computedState := E_FileExporterState.error;
			END_IF
		END_IF

	E_FileExporterState.done:
		IF NOT _execute THEN
			_computedState := E_FileExporterState.idle;
		END_IF
		THIS^.free();

	E_FileExporterState.error:
		// Retain the failure until export accepts a new batch.
END_CASE

currentState := _computedState;

IF currentState <= E_FileExporterState.serializing THEN _hFile := 0; END_IF
IF currentState = E_FileExporterState.done
	OR_ELSE currentState = E_FileExporterState.error THEN
	THIS^.free();
END_IF

_fileOpener(
	sNetId:='',
	sPathName:=THIS^._filepath,
	bExecute:=currentState = E_FileExporterState.opening,
	nMode:=FOPEN_MODEAPPEND OR FOPEN_MODETEXT,
	ePath:=PATH_GENERIC,
	tTimeout:=DEFAULT_ADS_TIMEOUT
);

_fileWriter(
	hFile:=_hFile,
	bExecute:=currentState = E_FileExporterState.writing,
	pWriteBuff:=_pString,
	cbWriteLen:=_len
);

_fileCloser(
	hFile:=_hFile,
	bExecute:=currentState = E_FileExporterState.closing
);

IF currentState = E_FileExporterState.error THEN
	tick := FALSE;
	failureReason := _failureReason;
END_IF
END_METHOD

END_FUNCTION_BLOCK

// ---- OTEL/LOGGING/SERIALIZATION/FUNCTION_BLOCKS/FB_LogRecordProtoJsonSerializer.TcPOU
FUNCTION_BLOCK FB_LogRecordProtoJsonSerializer EXTENDS FB_BaseProtoJsonSerializer

METHOD serializeLogRecord : BOOL
VAR_IN_OUT
	v: SJsonValue;
END_VAR
VAR_INPUT
	pLogRecord: POINTER TO FB_LogRecord;
END_VAR
VAR_OUTPUT
	failureReason: E_ProtoJsonSerializerFailureReason;
END_VAR
VAR
	_buf: T_MaxString;
	_obj: SJsonValue;
	_member: SJsonValue;
END_VAR
serializeLogRecord := FALSE;
failureReason := E_ProtoJsonSerializerFailureReason.NA;
IF v = 0 THEN
	failureReason := E_ProtoJsonSerializerFailureReason.JSON_VALUE_INVALID;
	RETURN;
END_IF
IF pLogRecord = 0 THEN
	failureReason := E_ProtoJsonSerializerFailureReason.LOG_RECORD_POINTER_NULL;
	RETURN;
END_IF

_obj := THIS^.parser.PushbackJsonValue(v, '{}');
IF _obj = 0 THEN
	failureReason := E_ProtoJsonSerializerFailureReason.JSON_OPERATION_FAILURE;
	RETURN;
END_IF

_buf := pLogRecord^.severityText;
_member := THIS^.parser.AddUintMember(_obj, 'severityNumber', TO_UDINT(pLogRecord^.severityNumber));
IF _member = 0 THEN failureReason := E_ProtoJsonSerializerFailureReason.JSON_OPERATION_FAILURE; RETURN; END_IF
_member := THIS^.parser.AddStringMember(_obj, 'severityText', _buf);
IF _member = 0 THEN failureReason := E_ProtoJsonSerializerFailureReason.JSON_OPERATION_FAILURE; RETURN; END_IF
IF NOT THIS^.serializeUint64Value(_obj, ADR('timeUnixNano'), pLogRecord^.timestamp, failureReason=>failureReason) THEN RETURN; END_IF

IF pLogRecord^.eventName <> 0 AND_THEN NOT THIS^.serializeStringValue(_obj, ADR('eventName'), pLogRecord^.eventName, failureReason=>failureReason) THEN RETURN; END_IF
IF pLogRecord^.traceId <> 0 AND_THEN NOT THIS^.serializeTraceIdValue(_obj, pLogRecord^.traceId, failureReason=>failureReason) THEN RETURN; END_IF
IF pLogRecord^.traceId <> 0 AND_THEN NOT THIS^.serializeUint32Value(_obj, ADR('flags'), TO_UDINT(pLogRecord^.flags), failureReason=>failureReason) THEN RETURN; END_IF
IF pLogRecord^.spanId <> 0 AND_THEN NOT THIS^.serializeSpanIdValue(_obj, pLogRecord^.spanId, failureReason=>failureReason) THEN RETURN; END_IF
IF pLogRecord^.body <> 0 AND_THEN NOT THIS^.serializeAnyValue(_obj, ADR('body'), pLogRecord^.body, failureReason=>failureReason) THEN RETURN; END_IF
IF pLogRecord^.attributes.count > 0 AND_THEN NOT THIS^.serializeKeyValues(_obj, ADR('attributes'), ADR(pLogRecord^.attributes), failureReason=>failureReason) THEN RETURN; END_IF
IF pLogRecord^.droppedAttributesCount > 0 AND_THEN NOT THIS^.serializeUint32Value(
	_obj,
	ADR('droppedAttributesCount'),
	pLogRecord^.droppedAttributesCount,
	failureReason=>failureReason
) THEN
	RETURN;
END_IF
serializeLogRecord := failureReason = E_ProtoJsonSerializerFailureReason.NA;
END_METHOD

(*
	Takes ownership of all supplied records. Popped records and records remaining in the
	queue are released on both success and failure.
*)
METHOD serializeLogsData : BOOL
VAR_IN_OUT
	logRecords: FB_LogRecordQueue;
END_VAR
VAR_OUTPUT
	failureReason: E_ProtoJsonSerializerFailureReason;
END_VAR
VAR
	_ownedRecordCount: UDINT;
	_pOwnedRecord: POINTER TO FB_LogRecord;
	_resourceLogs: SJsonValue;
	_resourceIdx: UDINT;
	_queueFailureReason: E_LogRecordQueueFailureReason;
END_VAR
serializeLogsData := FALSE;
failureReason := E_ProtoJsonSerializerFailureReason.NA;

// fail early if loop limit exceeded.
_ownedRecordCount := logRecords.count;
IF _ownedRecordCount > TcOtlp_GVL.MAX_LOOP_COUNT THEN
	logRecords.free();
	failureReason := E_ProtoJsonSerializerFailureReason.LOOP_LIMIT_EXCEEDED;
	RETURN;
END_IF

// start a new document in make the first entry an object i.e. "{}"
THIS^.jsonValue := THIS^.parser.NewDocument();
IF THIS^.jsonValue = 0 THEN
	logRecords.free();
	failureReason := E_ProtoJsonSerializerFailureReason.JSON_OPERATION_FAILURE;
	RETURN;
END_IF
THIS^.jsonValue := THIS^.parser.SetObject(THIS^.jsonValue);
IF THIS^.jsonValue = 0 THEN
	logRecords.free();
	failureReason := E_ProtoJsonSerializerFailureReason.JSON_OPERATION_FAILURE;
	RETURN;
END_IF

// start the resource logs block
_resourceLogs := THIS^.parser.AddArrayMember(THIS^.jsonValue, 'resourceLogs', 0);
IF _resourceLogs = 0 THEN
	logRecords.free();
	failureReason := E_ProtoJsonSerializerFailureReason.JSON_OPERATION_FAILURE;
	RETURN;
END_IF

_pOwnedRecord := 0;
IF _ownedRecordCount > 0 THEN
	FOR _resourceIdx := 1 TO _ownedRecordCount DO
		IF logRecords.count = 0 THEN EXIT; END_IF

		// pop the record to start the group
		IF NOT logRecords.pop(pValue:=_pOwnedRecord, failureReason=>_queueFailureReason) THEN
			failureReason := E_ProtoJsonSerializerFailureReason.QUEUE_POP_FAILURE;
			EXIT;
		END_IF
		IF _pOwnedRecord = 0 THEN
			failureReason := E_ProtoJsonSerializerFailureReason.LOG_RECORD_COLLECTION_INCONSISTENT;
			EXIT;
		END_IF

		// Recursively descend from LogsData into ResourceLogs and ScopeLogs.
		IF NOT THIS^.serializeResourceLogs(
			v:=_resourceLogs,
			logRecords:=logRecords,
			pLogRecord:=_pOwnedRecord,
			failureReason=>failureReason
		) THEN
			EXIT;
		END_IF
	END_FOR
END_IF

// clean up the last record if it's not cleaned up already
IF _pOwnedRecord <> 0 THEN
	_pOwnedRecord^.delete(pSelf:=_pOwnedRecord);
END_IF

// set flag if log records didn't all get consumed
IF logRecords.count > 0 THEN
	failureReason := E_ProtoJsonSerializerFailureReason.LOOP_LIMIT_EXCEEDED;
END_IF

// free all the memory and return status
logRecords.free();
serializeLogsData := failureReason = E_ProtoJsonSerializerFailureReason.NA;
END_METHOD

METHOD serializeResourceLogs : BOOL
VAR_IN_OUT
	v: SJsonValue;
	logRecords: FB_LogRecordQueue;
	pLogRecord: POINTER TO FB_LogRecord;
END_VAR
VAR_OUTPUT
	failureReason: E_ProtoJsonSerializerFailureReason;
END_VAR
VAR
	_resourceId: UDINT;
	_scopeLogs: SJsonValue;
	_pHeadRecord: POINTER TO FB_LogRecord;
	_scopeLimit: UDINT;
	_recordsToScan: UDINT;
	_scopeIdx: UDINT;
	_scanIdx: UDINT;
	_queueFailureReason: E_LogRecordQueueFailureReason;
END_VAR
serializeResourceLogs := FALSE;
failureReason := E_ProtoJsonSerializerFailureReason.NA;
IF v = 0 THEN
	failureReason := E_ProtoJsonSerializerFailureReason.JSON_VALUE_INVALID;
	RETURN;
END_IF
IF pLogRecord = 0 THEN
	failureReason := E_ProtoJsonSerializerFailureReason.LOG_RECORD_POINTER_NULL;
	RETURN;
END_IF

_resourceId := pLogRecord^.resource.id;
IF NOT THIS^.startNewResource(
	v:=v,
	pLogRecord:=pLogRecord,
	scopeLogs=>_scopeLogs,
	failureReason=>failureReason
) THEN
	RETURN;
END_IF

// Descend through each scope belonging to this resource. The queue remains
// the owner of every record until a matching record is popped.
_scopeLimit := logRecords.count + 1;
FOR _scopeIdx := 1 TO _scopeLimit DO
	IF NOT THIS^.serializeScopeLogs(
		v:=_scopeLogs,
		logRecords:=logRecords,
		pLogRecord:=pLogRecord,
		resourceId:=_resourceId,
		failureReason=>failureReason
	) THEN
		RETURN;
	END_IF

	// Find the first record for another scope of this resource. Rotating all
	// other records preserves their arrival order for later resource groups.
	_recordsToScan := logRecords.count;
	FOR _scanIdx := 1 TO _recordsToScan DO
		logRecords.reset();
		_pHeadRecord := logRecords.next();
		IF _pHeadRecord = 0 THEN
			failureReason := E_ProtoJsonSerializerFailureReason.LOG_RECORD_COLLECTION_INCONSISTENT;
			RETURN;
		END_IF
		IF pLogRecord = 0 AND_THEN _pHeadRecord^.resource.id = _resourceId THEN
			IF NOT logRecords.pop(pValue:=pLogRecord, failureReason=>_queueFailureReason) THEN
				failureReason := E_ProtoJsonSerializerFailureReason.QUEUE_POP_FAILURE;
				RETURN;
			END_IF
			IF pLogRecord = 0 THEN
				failureReason := E_ProtoJsonSerializerFailureReason.LOG_RECORD_COLLECTION_INCONSISTENT;
				RETURN;
			END_IF
		ELSIF NOT logRecords.rotate(failureReason=>_queueFailureReason) THEN
			failureReason := E_ProtoJsonSerializerFailureReason.QUEUE_ROTATE_FAILURE;
			RETURN;
		END_IF
	END_FOR

	IF pLogRecord = 0 THEN
		serializeResourceLogs := failureReason = E_ProtoJsonSerializerFailureReason.NA;
		RETURN;
	END_IF
END_FOR

failureReason := E_ProtoJsonSerializerFailureReason.LOOP_LIMIT_EXCEEDED;
END_METHOD

METHOD serializeScopeLogs : BOOL
VAR_IN_OUT
	v: SJsonValue;
	logRecords: FB_LogRecordQueue;
	pLogRecord: POINTER TO FB_LogRecord;
END_VAR
VAR_INPUT
	resourceId: UDINT;
END_VAR
VAR_OUTPUT
	failureReason: E_ProtoJsonSerializerFailureReason;
END_VAR
VAR
	_scopeName: T_MaxString;
	_serializedRecords: SJsonValue;
	_pHeadRecord: POINTER TO FB_LogRecord;
	_recordsToScan: UDINT;
	_scanIdx: UDINT;
	_queueFailureReason: E_LogRecordQueueFailureReason;
END_VAR
serializeScopeLogs := FALSE;
failureReason := E_ProtoJsonSerializerFailureReason.NA;
IF v = 0 THEN
	failureReason := E_ProtoJsonSerializerFailureReason.JSON_VALUE_INVALID;
	RETURN;
END_IF
IF pLogRecord = 0 THEN
	failureReason := E_ProtoJsonSerializerFailureReason.LOG_RECORD_POINTER_NULL;
	RETURN;
END_IF
IF pLogRecord^.resource.id <> resourceId THEN
	failureReason := E_ProtoJsonSerializerFailureReason.LOG_RECORD_COLLECTION_INCONSISTENT;
	RETURN;
END_IF

_scopeName := pLogRecord^.scope.name;
IF NOT THIS^.startNewScope(
	v:=v,
	pLogRecord:=pLogRecord,
	serializedRecords=>_serializedRecords,
	failureReason=>failureReason
) THEN
	RETURN;
END_IF

IF NOT THIS^.serializeLogRecord(_serializedRecords, pLogRecord, failureReason=>failureReason) THEN
	RETURN;
END_IF
pLogRecord^.delete(pSelf:=pLogRecord);

// Consume and release every remaining record in this resource/scope group.
_recordsToScan := logRecords.count;
FOR _scanIdx := 1 TO _recordsToScan DO
	logRecords.reset();
	_pHeadRecord := logRecords.next();
	IF _pHeadRecord = 0 THEN
		failureReason := E_ProtoJsonSerializerFailureReason.LOG_RECORD_COLLECTION_INCONSISTENT;
		RETURN;
	END_IF

	IF _pHeadRecord^.resource.id = resourceId AND_THEN _pHeadRecord^.scope.name = _scopeName THEN
		IF NOT logRecords.pop(pValue:=pLogRecord, failureReason=>_queueFailureReason) THEN
			failureReason := E_ProtoJsonSerializerFailureReason.QUEUE_POP_FAILURE;
			RETURN;
		END_IF
		IF pLogRecord = 0 THEN
			failureReason := E_ProtoJsonSerializerFailureReason.LOG_RECORD_COLLECTION_INCONSISTENT;
			RETURN;
		END_IF
		IF NOT THIS^.serializeLogRecord(_serializedRecords, pLogRecord, failureReason=>failureReason) THEN
			RETURN;
		END_IF
		pLogRecord^.delete(pSelf:=pLogRecord);
	ELSIF NOT logRecords.rotate(failureReason=>_queueFailureReason) THEN
		failureReason := E_ProtoJsonSerializerFailureReason.QUEUE_ROTATE_FAILURE;
		RETURN;
	END_IF
END_FOR

serializeScopeLogs := failureReason = E_ProtoJsonSerializerFailureReason.NA;
END_METHOD

METHOD startNewResource : BOOL
VAR_IN_OUT
	v: SJsonValue;
END_VAR
VAR_INPUT
	pLogRecord: POINTER TO FB_LogRecord;
END_VAR
VAR_OUTPUT
	scopeLogs: SJsonValue;
	failureReason: E_ProtoJsonSerializerFailureReason;
END_VAR
VAR
	_resourceObj: SJsonValue;
	_member: SJsonValue;
END_VAR
startNewResource := FALSE;
scopeLogs := 0;
failureReason := E_ProtoJsonSerializerFailureReason.NA;
IF v = 0 THEN
	failureReason := E_ProtoJsonSerializerFailureReason.JSON_VALUE_INVALID;
	RETURN;
END_IF
IF pLogRecord = 0 THEN
	failureReason := E_ProtoJsonSerializerFailureReason.LOG_RECORD_POINTER_NULL;
	RETURN;
END_IF

_resourceObj := THIS^.parser.PushbackJsonValue(v, '{}');
IF _resourceObj = 0 THEN
	failureReason := E_ProtoJsonSerializerFailureReason.JSON_OPERATION_FAILURE;
	RETURN;
END_IF
IF NOT THIS^._injectResource(_resourceObj, pLogRecord^.resource, failureReason=>failureReason) THEN
	RETURN;
END_IF
IF pLogRecord^.resource.schemaUrl <> '' THEN
	_member := THIS^.parser.AddStringMember(_resourceObj, 'schemaUrl', pLogRecord^.resource.schemaUrl);
	IF _member = 0 THEN
		failureReason := E_ProtoJsonSerializerFailureReason.JSON_OPERATION_FAILURE;
		RETURN;
	END_IF
END_IF
scopeLogs := THIS^.parser.AddArrayMember(_resourceObj, 'scopeLogs', 0);
IF scopeLogs = 0 THEN
	failureReason := E_ProtoJsonSerializerFailureReason.JSON_OPERATION_FAILURE;
	RETURN;
END_IF

startNewResource := failureReason = E_ProtoJsonSerializerFailureReason.NA;
END_METHOD

METHOD startNewScope : BOOL
VAR_IN_OUT
	v: SJsonValue;
END_VAR
VAR_INPUT
	pLogRecord: POINTER TO FB_LogRecord;
END_VAR
VAR_OUTPUT
	serializedRecords: SJsonValue;
	failureReason: E_ProtoJsonSerializerFailureReason;
END_VAR
VAR
	_scopeObj: SJsonValue;
	_member: SJsonValue;
END_VAR
startNewScope := FALSE;
serializedRecords := 0;
failureReason := E_ProtoJsonSerializerFailureReason.NA;
IF v = 0 THEN
	failureReason := E_ProtoJsonSerializerFailureReason.JSON_VALUE_INVALID;
	RETURN;
END_IF
IF pLogRecord = 0 THEN
	failureReason := E_ProtoJsonSerializerFailureReason.LOG_RECORD_POINTER_NULL;
	RETURN;
END_IF

_scopeObj := THIS^.parser.PushbackJsonValue(v, '{}');
IF _scopeObj = 0 THEN
	failureReason := E_ProtoJsonSerializerFailureReason.JSON_OPERATION_FAILURE;
	RETURN;
END_IF
IF NOT THIS^._injectInstrumentationScope(_scopeObj, pLogRecord^.scope, failureReason=>failureReason) THEN
	RETURN;
END_IF
IF pLogRecord^.scope.schemaUrl <> '' THEN
	_member := THIS^.parser.AddStringMember(_scopeObj, 'schemaUrl', pLogRecord^.scope.schemaUrl);
	IF _member = 0 THEN
		failureReason := E_ProtoJsonSerializerFailureReason.JSON_OPERATION_FAILURE;
		RETURN;
	END_IF
END_IF
serializedRecords := THIS^.parser.AddArrayMember(_scopeObj, 'logRecords', 0);
IF serializedRecords = 0 THEN
	failureReason := E_ProtoJsonSerializerFailureReason.JSON_OPERATION_FAILURE;
	RETURN;
END_IF

startNewScope := failureReason = E_ProtoJsonSerializerFailureReason.NA;
END_METHOD

END_FUNCTION_BLOCK

// ---- OTEL/SERIALIZATION/FUNCTION_BLOCKS/FB_BaseProtoJsonSerializer.TcPOU
FUNCTION_BLOCK FB_BaseProtoJsonSerializer

VAR_OUTPUT
	parser: FB_JsonDynDomParser;
	jsonValue: SJsonValue;
END_VAR

METHOD _injectInstrumentationScope : BOOL
VAR_IN_OUT
	v: SJsonValue;
	instrumentationScope: FB_InstrumentationScope;
END_VAR
VAR_OUTPUT
	failureReason: E_ProtoJsonSerializerFailureReason;
END_VAR
VAR
	_obj: SJsonValue;
	_member: SJsonValue;
END_VAR
_injectInstrumentationScope := FALSE;
failureReason := E_ProtoJsonSerializerFailureReason.NA;
IF v = 0 THEN
	failureReason := E_ProtoJsonSerializerFailureReason.JSON_VALUE_INVALID;
	RETURN;
END_IF

_obj := THIS^.parser.AddObjectMember(v, 'scope');
IF _obj = 0 THEN
	failureReason := E_ProtoJsonSerializerFailureReason.JSON_OPERATION_FAILURE;
	RETURN;
END_IF
_member := THIS^.parser.AddStringMember(_obj, 'name', instrumentationScope.name);
IF _member = 0 THEN
	failureReason := E_ProtoJsonSerializerFailureReason.JSON_OPERATION_FAILURE;
	RETURN;
END_IF
_member := THIS^.parser.AddStringMember(_obj, 'version', instrumentationScope.version);
IF _member = 0 THEN
	failureReason := E_ProtoJsonSerializerFailureReason.JSON_OPERATION_FAILURE;
	RETURN;
END_IF
IF instrumentationScope.attributes.count > 0 AND_THEN NOT THIS^.serializeKeyValues(
	v:=_obj,
	pKey:=ADR('attributes'),
	pValues:=ADR(instrumentationScope.attributes),
	failureReason=>failureReason
) THEN
	RETURN;
END_IF
IF instrumentationScope.attributes.count > 0 OR instrumentationScope.droppedAttributesCount > 0 THEN
	IF NOT THIS^.serializeUint32Value(
		v:=_obj,
		pKey:=ADR('droppedAttributesCount'),
		val:=instrumentationScope.droppedAttributesCount,
		failureReason=>failureReason
	) THEN
		RETURN;
	END_IF
END_IF
_injectInstrumentationScope := failureReason = E_ProtoJsonSerializerFailureReason.NA;
END_METHOD

METHOD _injectResource : BOOL
VAR_IN_OUT
	v: SJsonValue;
	resource: FB_Resource;
END_VAR
VAR_OUTPUT
	failureReason: E_ProtoJsonSerializerFailureReason;
END_VAR
VAR
	_obj: SJsonValue;
END_VAR
_injectResource := FALSE;
failureReason := E_ProtoJsonSerializerFailureReason.NA;
IF v = 0 THEN
	failureReason := E_ProtoJsonSerializerFailureReason.JSON_VALUE_INVALID;
	RETURN;
END_IF

_obj := THIS^.parser.AddObjectMember(v, 'resource');
IF _obj = 0 THEN
	failureReason := E_ProtoJsonSerializerFailureReason.JSON_OPERATION_FAILURE;
	RETURN;
END_IF
IF resource.attributes.count > 0 AND_THEN NOT THIS^.serializeKeyValues(
	v:=_obj,
	pKey:=ADR('attributes'),
	pValues:=ADR(resource.attributes),
	failureReason=>failureReason
) THEN
	RETURN;
END_IF
IF resource.droppedAttributesCount > 0 AND_THEN NOT THIS^.serializeUint32Value(
	v:=_obj,
	pKey:=ADR('droppedAttributesCount'),
	val:=resource.droppedAttributesCount,
	failureReason=>failureReason
) THEN
	RETURN;
END_IF
_injectResource := failureReason = E_ProtoJsonSerializerFailureReason.NA;
END_METHOD

METHOD _serializeBytes : BOOL
VAR_INPUT
	pBytes: POINTER TO BYTE;
	nBytes: UDINT := 0;
	pStr: POINTER TO STRING;
	len: UDINT;
	encoding: E_BytesEncoding;
END_VAR
VAR_OUTPUT
	failureReason: E_ProtoJsonSerializerFailureReason;
END_VAR
VAR
	_idx: UDINT;
	_nibble: BYTE;
	_requiredLen: UDINT;
END_VAR
_serializeBytes := FALSE;
failureReason := E_ProtoJsonSerializerFailureReason.NA;
IF pBytes = 0 THEN
	failureReason := E_ProtoJsonSerializerFailureReason.BYTES_POINTER_NULL;
	RETURN;
END_IF
IF nBytes = 0 THEN
	failureReason := E_ProtoJsonSerializerFailureReason.BYTE_COUNT_ZERO;
	RETURN;
END_IF
IF pStr = 0 THEN
	failureReason := E_ProtoJsonSerializerFailureReason.STRING_POINTER_NULL;
	RETURN;
END_IF

_requiredLen := nBytes * 2;
IF len <= _requiredLen THEN
	failureReason := E_ProtoJsonSerializerFailureReason.STRING_BUFFER_TOO_SMALL;
	RETURN;
END_IF
IF encoding <> E_BytesEncoding.hex THEN
	failureReason := E_ProtoJsonSerializerFailureReason.UNSUPPORTED_BYTES_ENCODING;
	RETURN;
END_IF

pStr^ := '';
FOR _idx := 0 TO nBytes - 1 DO
	_nibble := SHR(pBytes[_idx], 4) AND 16#0F;
	pStr^[(_idx * 2)] := SEL(_nibble < 10, _nibble + 16#37, _nibble + 16#30);
	_nibble := pBytes[_idx] AND 16#0F;
	pStr^[(_idx * 2) + 1] := SEL(_nibble < 10, _nibble + 16#37, _nibble + 16#30);
END_FOR
pStr^[_requiredLen] := 0;
_serializeBytes :=failureReason = E_ProtoJsonSerializerFailureReason.NA;
END_METHOD

METHOD serializeAnyValue : BOOL
VAR_IN_OUT
	v: SJsonValue;
END_VAR
VAR_INPUT
	pKey: POINTER TO STRING;
	pVal: POINTER TO FB_AnyValue;
END_VAR
VAR_OUTPUT
	failureReason: E_ProtoJsonSerializerFailureReason;
END_VAR
VAR
	_v: SJsonValue;
	_pNumber: POINTER TO FB_Number;
	_pSInt: POINTER TO SINT;
	_pInt: POINTER TO INT;
	_pDInt: POINTER TO DINT;
	_pLInt: POINTER TO LINT;
	_pUSInt: POINTER TO USINT;
	_pUInt: POINTER TO UINT;
	_pUDInt: POINTER TO UDINT;
	_pULInt: POINTER TO ULINT;
	_pReal: POINTER TO REAL;
	_pLReal: POINTER TO LREAL;
END_VAR
serializeAnyValue := FALSE;
failureReason := E_ProtoJsonSerializerFailureReason.NA;
IF v = 0 THEN
	failureReason := E_ProtoJsonSerializerFailureReason.JSON_VALUE_INVALID;
	RETURN;
END_IF
IF pKey = 0 THEN
	failureReason := E_ProtoJsonSerializerFailureReason.KEY_POINTER_NULL;
	RETURN;
END_IF
IF pVal = 0 THEN
	failureReason := E_ProtoJsonSerializerFailureReason.VALUE_POINTER_NULL;
	RETURN;
END_IF

_v := THIS^.parser.AddObjectMember(v, pKey^);
IF _v = 0 THEN
	failureReason := E_ProtoJsonSerializerFailureReason.JSON_OPERATION_FAILURE;
	RETURN;
END_IF

CASE pVal^.eType OF
	E_ValueType.E_String:
		serializeAnyValue := THIS^.serializeStringValue(
			v:=_v,
			pKey:=ADR('stringValue'),
			pVal:=pVal,
			failureReason=>failureReason
		);
	E_ValueType.E_Number:
		_pNumber := pVal;
		IF _pNumber^.value.pValue = 0 THEN
			failureReason := E_ProtoJsonSerializerFailureReason.NUMBER_VALUE_POINTER_NULL;
			RETURN;
		END_IF
		CASE _pNumber^.value.TypeClass OF
			__SYSTEM.TYPE_CLASS.TYPE_SINT:
				_pSInt := _pNumber^.value.pValue;
				serializeAnyValue := THIS^.serializeInt64Value(_v, ADR('intValue'), SINT_TO_LINT(_pSInt^), failureReason=>failureReason);
			__SYSTEM.TYPE_CLASS.TYPE_INT:
				_pInt := _pNumber^.value.pValue;
				serializeAnyValue := THIS^.serializeInt64Value(_v, ADR('intValue'), INT_TO_LINT(_pInt^), failureReason=>failureReason);
			__SYSTEM.TYPE_CLASS.TYPE_DINT:
				_pDInt := _pNumber^.value.pValue;
				serializeAnyValue := THIS^.serializeInt64Value(_v, ADR('intValue'), DINT_TO_LINT(_pDInt^), failureReason=>failureReason);
			__SYSTEM.TYPE_CLASS.TYPE_LINT:
				_pLInt := _pNumber^.value.pValue;
				serializeAnyValue := THIS^.serializeInt64Value(_v, ADR('intValue'), _pLInt^, failureReason=>failureReason);
			__SYSTEM.TYPE_CLASS.TYPE_USINT:
				_pUSInt := _pNumber^.value.pValue;
				serializeAnyValue := THIS^.serializeUint64Value(_v, ADR('intValue'), USINT_TO_ULINT(_pUSInt^), failureReason=>failureReason);
			__SYSTEM.TYPE_CLASS.TYPE_UINT:
				_pUInt := _pNumber^.value.pValue;
				serializeAnyValue := THIS^.serializeUint64Value(_v, ADR('intValue'), UINT_TO_ULINT(_pUInt^), failureReason=>failureReason);
			__SYSTEM.TYPE_CLASS.TYPE_UDINT:
				_pUDInt := _pNumber^.value.pValue;
				serializeAnyValue := THIS^.serializeUint64Value(_v, ADR('intValue'), UDINT_TO_ULINT(_pUDInt^), failureReason=>failureReason);
			__SYSTEM.TYPE_CLASS.TYPE_ULINT:
				_pULInt := _pNumber^.value.pValue;
				serializeAnyValue := THIS^.serializeUint64Value(_v, ADR('intValue'), _pULInt^, failureReason=>failureReason);
			__SYSTEM.TYPE_CLASS.TYPE_REAL:
				_pReal := _pNumber^.value.pValue;
				serializeAnyValue := THIS^.serializeDoubleValue(_v, ADR('doubleValue'), REAL_TO_LREAL(_pReal^), failureReason=>failureReason);
			__SYSTEM.TYPE_CLASS.TYPE_LREAL:
				_pLReal := _pNumber^.value.pValue;
				serializeAnyValue := THIS^.serializeDoubleValue(_v, ADR('doubleValue'), _pLReal^, failureReason=>failureReason);
			ELSE
				failureReason := E_ProtoJsonSerializerFailureReason.UNSUPPORTED_NUMBER_TYPE;
		END_CASE
	ELSE
		failureReason := E_ProtoJsonSerializerFailureReason.UNSUPPORTED_VALUE_TYPE;
END_CASE
END_METHOD

METHOD serializeDoubleValue : BOOL
VAR_IN_OUT
	v: SJsonValue;
END_VAR
VAR_INPUT
	pKey: POINTER TO STRING;
	val: LREAL;
END_VAR
VAR_OUTPUT
	failureReason: E_ProtoJsonSerializerFailureReason;
END_VAR
VAR
	_bits: LWORD;
	_member: SJsonValue;
END_VAR
serializeDoubleValue := FALSE;
failureReason := E_ProtoJsonSerializerFailureReason.NA;
IF v = 0 THEN failureReason := E_ProtoJsonSerializerFailureReason.JSON_VALUE_INVALID; RETURN; END_IF
IF pKey = 0 THEN failureReason := E_ProtoJsonSerializerFailureReason.KEY_POINTER_NULL; RETURN; END_IF

MEMCPY(ADR(_bits), ADR(val), SIZEOF(_bits));
IF (_bits AND LWORD#16#7FF0000000000000) = LWORD#16#7FF0000000000000 THEN
	IF (_bits AND LWORD#16#000FFFFFFFFFFFFF) <> 0 THEN
		_member := THIS^.parser.AddStringMember(v, pKey^, 'NaN');
	ELSIF (_bits AND LWORD#16#8000000000000000) <> 0 THEN
		_member := THIS^.parser.AddStringMember(v, pKey^, '-Infinity');
	ELSE
		_member := THIS^.parser.AddStringMember(v, pKey^, 'Infinity');
	END_IF
ELSE
	_member := THIS^.parser.AddDoubleMember(v, pKey^, val);
END_IF
IF _member = 0 THEN failureReason := E_ProtoJsonSerializerFailureReason.JSON_OPERATION_FAILURE; RETURN; END_IF
serializeDoubleValue := failureReason = E_ProtoJsonSerializerFailureReason.NA;
END_METHOD

METHOD serializeFloatValue : BOOL
VAR_IN_OUT
	v: SJsonValue;
END_VAR
VAR_INPUT
	pKey: POINTER TO STRING;
	val: REAL;
END_VAR
VAR_OUTPUT
	failureReason: E_ProtoJsonSerializerFailureReason;
END_VAR
VAR
	_bits: DWORD;
	_member: SJsonValue;
END_VAR
serializeFloatValue := FALSE;
failureReason := E_ProtoJsonSerializerFailureReason.NA;
IF v = 0 THEN failureReason := E_ProtoJsonSerializerFailureReason.JSON_VALUE_INVALID; RETURN; END_IF
IF pKey = 0 THEN failureReason := E_ProtoJsonSerializerFailureReason.KEY_POINTER_NULL; RETURN; END_IF

MEMCPY(ADR(_bits), ADR(val), SIZEOF(_bits));
IF (_bits AND DWORD#16#7F800000) = DWORD#16#7F800000 THEN
	IF (_bits AND DWORD#16#007FFFFF) <> 0 THEN
		_member := THIS^.parser.AddStringMember(v, pKey^, 'NaN');
	ELSIF (_bits AND DWORD#16#80000000) <> 0 THEN
		_member := THIS^.parser.AddStringMember(v, pKey^, '-Infinity');
	ELSE
		_member := THIS^.parser.AddStringMember(v, pKey^, 'Infinity');
	END_IF
ELSE
	_member := THIS^.parser.AddDoubleMember(v, pKey^, REAL_TO_LREAL(val));
END_IF
IF _member = 0 THEN failureReason := E_ProtoJsonSerializerFailureReason.JSON_OPERATION_FAILURE; RETURN; END_IF
serializeFloatValue := failureReason = E_ProtoJsonSerializerFailureReason.NA;
END_METHOD

METHOD serializeInt32Value : BOOL
VAR_IN_OUT
	v: SJsonValue;
END_VAR
VAR_INPUT
	pKey: POINTER TO STRING;
	val: DINT;
END_VAR
VAR_OUTPUT
	failureReason: E_ProtoJsonSerializerFailureReason;
END_VAR
VAR
	_member: SJsonValue;
END_VAR
serializeInt32Value := FALSE;
failureReason := E_ProtoJsonSerializerFailureReason.NA;
IF v = 0 THEN failureReason := E_ProtoJsonSerializerFailureReason.JSON_VALUE_INVALID; RETURN; END_IF
IF pKey = 0 THEN failureReason := E_ProtoJsonSerializerFailureReason.KEY_POINTER_NULL; RETURN; END_IF
_member := THIS^.parser.AddIntMember(v, pKey^, val);
IF _member = 0 THEN failureReason := E_ProtoJsonSerializerFailureReason.JSON_OPERATION_FAILURE; RETURN; END_IF
serializeInt32Value := failureReason = E_ProtoJsonSerializerFailureReason.NA;
END_METHOD

METHOD serializeInt64Value : BOOL
VAR_IN_OUT
	v: SJsonValue;
END_VAR
VAR_INPUT
	pKey: POINTER TO STRING;
	val: LINT;
END_VAR
VAR_OUTPUT
	failureReason: E_ProtoJsonSerializerFailureReason;
END_VAR
VAR
	_buf: STRING(20);
	_member: SJsonValue;
END_VAR
serializeInt64Value := FALSE;
failureReason := E_ProtoJsonSerializerFailureReason.NA;
IF v = 0 THEN failureReason := E_ProtoJsonSerializerFailureReason.JSON_VALUE_INVALID; RETURN; END_IF
IF pKey = 0 THEN failureReason := E_ProtoJsonSerializerFailureReason.KEY_POINTER_NULL; RETURN; END_IF
_buf := LINT_TO_STRING(val);
_member := THIS^.parser.AddStringMember(v, pKey^, _buf);
IF _member = 0 THEN failureReason := E_ProtoJsonSerializerFailureReason.JSON_OPERATION_FAILURE; RETURN; END_IF
serializeInt64Value := failureReason = E_ProtoJsonSerializerFailureReason.NA;
END_METHOD

METHOD serializeKeyValue : BOOL
VAR_IN_OUT
	v: SJsonValue;
END_VAR
VAR_INPUT
	pVal: POINTER TO FB_KeyValue;
END_VAR
VAR_OUTPUT
	failureReason: E_ProtoJsonSerializerFailureReason;
END_VAR
VAR
	_member: SJsonValue;
END_VAR
serializeKeyValue := FALSE;
failureReason := E_ProtoJsonSerializerFailureReason.NA;
IF v = 0 THEN failureReason := E_ProtoJsonSerializerFailureReason.JSON_VALUE_INVALID; RETURN; END_IF
IF pVal = 0 OR_ELSE pVal^.pVal = 0 THEN failureReason := E_ProtoJsonSerializerFailureReason.VALUE_POINTER_NULL; RETURN; END_IF
IF pVal^.pKey = 0 THEN failureReason := E_ProtoJsonSerializerFailureReason.KEY_POINTER_NULL; RETURN; END_IF
_member := THIS^.parser.AddStringMember(v, 'key', pVal^.pKey^);
IF _member = 0 THEN failureReason := E_ProtoJsonSerializerFailureReason.JSON_OPERATION_FAILURE; RETURN; END_IF
serializeKeyValue := THIS^.serializeAnyValue(v, ADR('value'), pVal^.pVal, failureReason=>failureReason);
END_METHOD

METHOD serializeKeyValues : BOOL
VAR_IN_OUT
	v: SJsonValue;
END_VAR
VAR_INPUT
	pKey: POINTER TO STRING;
	pValues: POINTER TO FB_Attributes;
END_VAR
VAR_OUTPUT
	failureReason: E_ProtoJsonSerializerFailureReason;
END_VAR
VAR
	_idx: UDINT;
	_arr: SJsonValue;
	_obj: SJsonValue;
	_pValue: POINTER TO FB_KeyValue;
END_VAR
serializeKeyValues := FALSE;
failureReason := E_ProtoJsonSerializerFailureReason.NA;
IF v = 0 THEN failureReason := E_ProtoJsonSerializerFailureReason.JSON_VALUE_INVALID; RETURN; END_IF
IF pKey = 0 THEN failureReason := E_ProtoJsonSerializerFailureReason.KEY_POINTER_NULL; RETURN; END_IF
IF pValues = 0 THEN failureReason := E_ProtoJsonSerializerFailureReason.VALUE_POINTER_NULL; RETURN; END_IF
IF pValues^.count = 0 THEN serializeKeyValues := failureReason = E_ProtoJsonSerializerFailureReason.NA; RETURN; END_IF
IF pValues^.count > pValues^.maxCount OR_ELSE pValues^.count > TcOtlp_GVL.MAX_LOOP_COUNT THEN
	failureReason := E_ProtoJsonSerializerFailureReason.LOOP_LIMIT_EXCEEDED;
	RETURN;
END_IF

_arr := THIS^.parser.AddArrayMember(v, pKey^, 0);
IF _arr = 0 THEN failureReason := E_ProtoJsonSerializerFailureReason.JSON_OPERATION_FAILURE; RETURN; END_IF
pValues^.reset();
FOR _idx := 1 TO pValues^.count DO
	_pValue := pValues^.next();
	IF _pValue = 0 THEN
		pValues^.reset();
		failureReason := E_ProtoJsonSerializerFailureReason.ATTRIBUTE_COLLECTION_INCONSISTENT;
		RETURN;
	END_IF
	_obj := THIS^.parser.PushbackJsonValue(_arr, '{}');
	IF _obj = 0 THEN
		pValues^.reset();
		failureReason := E_ProtoJsonSerializerFailureReason.JSON_OPERATION_FAILURE;
		RETURN;
	END_IF
	IF NOT THIS^.serializeKeyValue(_obj, _pValue, failureReason=>failureReason) THEN
		pValues^.reset();
		RETURN;
	END_IF
END_FOR
pValues^.reset();
serializeKeyValues := failureReason = E_ProtoJsonSerializerFailureReason.NA;
END_METHOD

METHOD serializeNumberValue : BOOL
VAR_IN_OUT
	v: SJsonValue;
END_VAR
VAR_INPUT
	pKey: POINTER TO STRING;
	val: ANY_NUM;
END_VAR
VAR_OUTPUT
	failureReason: E_ProtoJsonSerializerFailureReason;
END_VAR
VAR
	_pSInt: POINTER TO SINT;
	_pInt: POINTER TO INT;
	_pDInt: POINTER TO DINT;
	_pLInt: POINTER TO LINT;
	_pUSInt: POINTER TO USINT;
	_pUInt: POINTER TO UINT;
	_pUDInt: POINTER TO UDINT;
	_pULInt: POINTER TO ULINT;
	_pReal: POINTER TO REAL;
	_pLReal: POINTER TO LREAL;
END_VAR
serializeNumberValue := FALSE;
failureReason := E_ProtoJsonSerializerFailureReason.NA;
IF v = 0 THEN failureReason := E_ProtoJsonSerializerFailureReason.JSON_VALUE_INVALID; RETURN; END_IF
IF pKey = 0 THEN failureReason := E_ProtoJsonSerializerFailureReason.KEY_POINTER_NULL; RETURN; END_IF
IF val.pValue = 0 THEN failureReason := E_ProtoJsonSerializerFailureReason.NUMBER_VALUE_POINTER_NULL; RETURN; END_IF

CASE val.TypeClass OF
	__SYSTEM.TYPE_CLASS.TYPE_SINT:
		_pSInt := val.pValue;
		serializeNumberValue := THIS^.serializeInt32Value(v, pKey, SINT_TO_DINT(_pSInt^), failureReason=>failureReason);
	__SYSTEM.TYPE_CLASS.TYPE_INT:
		_pInt := val.pValue;
		serializeNumberValue := THIS^.serializeInt32Value(v, pKey, INT_TO_DINT(_pInt^), failureReason=>failureReason);
	__SYSTEM.TYPE_CLASS.TYPE_DINT:
		_pDInt := val.pValue;
		serializeNumberValue := THIS^.serializeInt32Value(v, pKey, _pDInt^, failureReason=>failureReason);
	__SYSTEM.TYPE_CLASS.TYPE_LINT:
		_pLInt := val.pValue;
		serializeNumberValue := THIS^.serializeInt64Value(v, pKey, _pLInt^, failureReason=>failureReason);
	__SYSTEM.TYPE_CLASS.TYPE_USINT:
		_pUSInt := val.pValue;
		serializeNumberValue := THIS^.serializeUint32Value(v, pKey, USINT_TO_UDINT(_pUSInt^), failureReason=>failureReason);
	__SYSTEM.TYPE_CLASS.TYPE_UINT:
		_pUInt := val.pValue;
		serializeNumberValue := THIS^.serializeUint32Value(v, pKey, UINT_TO_UDINT(_pUInt^), failureReason=>failureReason);
	__SYSTEM.TYPE_CLASS.TYPE_UDINT:
		_pUDInt := val.pValue;
		serializeNumberValue := THIS^.serializeUint32Value(v, pKey, _pUDInt^, failureReason=>failureReason);
	__SYSTEM.TYPE_CLASS.TYPE_ULINT:
		_pULInt := val.pValue;
		serializeNumberValue := THIS^.serializeUint64Value(v, pKey, _pULInt^, failureReason=>failureReason);
	__SYSTEM.TYPE_CLASS.TYPE_REAL:
		_pReal := val.pValue;
		serializeNumberValue := THIS^.serializeFloatValue(v, pKey, _pReal^, failureReason=>failureReason);
	__SYSTEM.TYPE_CLASS.TYPE_LREAL:
		_pLReal := val.pValue;
		serializeNumberValue := THIS^.serializeDoubleValue(v, pKey, _pLReal^, failureReason=>failureReason);
	ELSE
		failureReason := E_ProtoJsonSerializerFailureReason.UNSUPPORTED_NUMBER_TYPE;
END_CASE
END_METHOD

METHOD serializeSpanIdValue : BOOL
VAR_IN_OUT
	v: SJsonValue;
END_VAR
VAR_INPUT
	pVal: POINTER TO FB_SpanId;
END_VAR
VAR_OUTPUT
	failureReason: E_ProtoJsonSerializerFailureReason;
END_VAR
VAR
	_encodedStr: STRING(16);
	_member: SJsonValue;
END_VAR
serializeSpanIdValue := FALSE;
failureReason := E_ProtoJsonSerializerFailureReason.NA;
IF v = 0 THEN failureReason := E_ProtoJsonSerializerFailureReason.JSON_VALUE_INVALID; RETURN; END_IF
IF pVal = 0 THEN failureReason := E_ProtoJsonSerializerFailureReason.VALUE_POINTER_NULL; RETURN; END_IF
IF NOT THIS^._serializeBytes(ADR(pVal^.bytes), SIZEOF(pVal^.bytes), ADR(_encodedStr), SIZEOF(_encodedStr), E_BytesEncoding.hex, failureReason=>failureReason) THEN RETURN; END_IF
_member := THIS^.parser.AddStringMember(v, 'spanId', _encodedStr);
IF _member = 0 THEN failureReason := E_ProtoJsonSerializerFailureReason.JSON_OPERATION_FAILURE; RETURN; END_IF
serializeSpanIdValue := failureReason = E_ProtoJsonSerializerFailureReason.NA;
END_METHOD

METHOD serializeStringValue : BOOL
VAR_IN_OUT
	v: SJsonValue;
END_VAR
VAR_INPUT
	pKey: POINTER TO STRING;
	pVal: POINTER TO FB_String;
END_VAR
VAR_OUTPUT
	failureReason: E_ProtoJsonSerializerFailureReason;
END_VAR
VAR
	_member: SJsonValue;
END_VAR
serializeStringValue := FALSE;
failureReason := E_ProtoJsonSerializerFailureReason.NA;
IF v = 0 THEN failureReason := E_ProtoJsonSerializerFailureReason.JSON_VALUE_INVALID; RETURN; END_IF
IF pKey = 0 THEN failureReason := E_ProtoJsonSerializerFailureReason.KEY_POINTER_NULL; RETURN; END_IF
IF pVal = 0 THEN failureReason := E_ProtoJsonSerializerFailureReason.VALUE_POINTER_NULL; RETURN; END_IF
IF pVal^.pString = 0 THEN failureReason := E_ProtoJsonSerializerFailureReason.STRING_POINTER_NULL; RETURN; END_IF
_member := THIS^.parser.AddStringMember(v, pKey^, pVal^.pString^);
IF _member = 0 THEN failureReason := E_ProtoJsonSerializerFailureReason.JSON_OPERATION_FAILURE; RETURN; END_IF
serializeStringValue := failureReason = E_ProtoJsonSerializerFailureReason.NA;
END_METHOD

METHOD serializeTraceIdValue : BOOL
VAR_IN_OUT
	v: SJsonValue;
END_VAR
VAR_INPUT
	pVal: POINTER TO FB_TraceId;
END_VAR
VAR_OUTPUT
	failureReason: E_ProtoJsonSerializerFailureReason;
END_VAR
VAR
	_encodedStr: STRING(32);
	_member: SJsonValue;
END_VAR
serializeTraceIdValue := FALSE;
failureReason := E_ProtoJsonSerializerFailureReason.NA;
IF v = 0 THEN failureReason := E_ProtoJsonSerializerFailureReason.JSON_VALUE_INVALID; RETURN; END_IF
IF pVal = 0 THEN failureReason := E_ProtoJsonSerializerFailureReason.VALUE_POINTER_NULL; RETURN; END_IF
IF NOT THIS^._serializeBytes(ADR(pVal^.bytes), SIZEOF(pVal^.bytes), ADR(_encodedStr), SIZEOF(_encodedStr), E_BytesEncoding.hex, failureReason=>failureReason) THEN RETURN; END_IF
_member := THIS^.parser.AddStringMember(v, 'traceId', _encodedStr);
IF _member = 0 THEN failureReason := E_ProtoJsonSerializerFailureReason.JSON_OPERATION_FAILURE; RETURN; END_IF
serializeTraceIdValue := failureReason = E_ProtoJsonSerializerFailureReason.NA;
END_METHOD

METHOD serializeUint32Value : BOOL
VAR_IN_OUT
	v: SJsonValue;
END_VAR
VAR_INPUT
	pKey: POINTER TO STRING;
	val: UDINT;
END_VAR
VAR_OUTPUT
	failureReason: E_ProtoJsonSerializerFailureReason;
END_VAR
VAR
	_member: SJsonValue;
END_VAR
serializeUint32Value := FALSE;
failureReason := E_ProtoJsonSerializerFailureReason.NA;
IF v = 0 THEN failureReason := E_ProtoJsonSerializerFailureReason.JSON_VALUE_INVALID; RETURN; END_IF
IF pKey = 0 THEN failureReason := E_ProtoJsonSerializerFailureReason.KEY_POINTER_NULL; RETURN; END_IF
_member := THIS^.parser.AddUintMember(v, pKey^, val);
IF _member = 0 THEN failureReason := E_ProtoJsonSerializerFailureReason.JSON_OPERATION_FAILURE; RETURN; END_IF
serializeUint32Value := failureReason = E_ProtoJsonSerializerFailureReason.NA;
END_METHOD

METHOD serializeUint64Value : BOOL
VAR_IN_OUT
	v: SJsonValue;
END_VAR
VAR_INPUT
	pKey: POINTER TO STRING;
	val: ULINT;
END_VAR
VAR_OUTPUT
	failureReason: E_ProtoJsonSerializerFailureReason;
END_VAR
VAR
	_buf: STRING(20);
	_member: SJsonValue;
END_VAR
serializeUint64Value := FALSE;
failureReason := E_ProtoJsonSerializerFailureReason.NA;
IF v = 0 THEN failureReason := E_ProtoJsonSerializerFailureReason.JSON_VALUE_INVALID; RETURN; END_IF
IF pKey = 0 THEN failureReason := E_ProtoJsonSerializerFailureReason.KEY_POINTER_NULL; RETURN; END_IF
_buf := ULINT_TO_STRING(val);
_member := THIS^.parser.AddStringMember(v, pKey^, _buf);
IF _member = 0 THEN failureReason := E_ProtoJsonSerializerFailureReason.JSON_OPERATION_FAILURE; RETURN; END_IF
serializeUint64Value := failureReason = E_ProtoJsonSerializerFailureReason.NA;
END_METHOD

END_FUNCTION_BLOCK

// ---- OTEL/LOGGING/EXPORTING/FUNCTION_BLOCKS/FB_LogRecordExporter_HTTP.TcPOU
FUNCTION_BLOCK FB_LogRecordExporter_HTTP EXTENDS FB_LogRecordExporter_Base
VAR_OUTPUT
	currentState: E_HttpExporterState;
	statusCode: UINT;  // the HTTP status code received for the last completed request
END_VAR

VAR
	_execute: BOOL;
	_urlParsed: BOOL;
	_endpoint: ST_HttpEndpoint;
	_len: UDINT;
	_execRTrig: R_TRIG;
	_pString: POINTER TO STRING;
	_jsonVal: SJsonValue;
	_computedState: E_HttpExporterState;
	_failureReason: E_LogRecordExporterFailureReason;
	_serializationFailureReason: E_ProtoJsonSerializerFailureReason;
	_serializer: FB_LogRecordProtoJsonSerializer;
	_client: FB_IotHttpClient;
	_request: FB_IotHttpRequest;
	_header: FB_IotHttpHeaderFieldMap;
END_VAR

THIS^.tick(failureReason=>THIS^._callFailureReason);

METHOD export: BOOL
VAR_IN_OUT
	logRecords: FB_LogRecordQueue;
END_VAR
VAR_INPUT
	count: UDINT;
END_VAR
VAR_OUTPUT
	failureReason: E_LogRecordExporterFailureReason;
END_VAR
// Prepare a completed exporter to accept the next batch immediately.
IF THIS^.currentState = E_HttpExporterState.done OR THIS^.currentState = E_HttpExporterState.error THEN
	THIS^.currentState := E_HttpExporterState.idle;
	THIS^._computedState := E_HttpExporterState.idle;
END_IF
export := SUPER^.export(
	logRecords:=logRecords,
	count:=count,
	failureReason=>failureReason
);
IF export THEN
	THIS^._failureReason := E_LogRecordExporterFailureReason.NA;
	THIS^._serializationFailureReason := E_ProtoJsonSerializerFailureReason.NA;
END_IF
END_METHOD

(*
	Releases a payload buffer that is still in flight. The FB_IotHttpRequest reading it is
	destroyed with this instance, so nothing uses the buffer afterwards. TwinCAT then
	runs FB_LogRecordExporter_Base.FB_Exit, which releases the queued records.
*)
METHOD FB_Exit : BOOL
VAR_INPUT
	bInCopyCode: BOOL;  // TRUE: the instance is being copied during an online change
END_VAR
// during an online change the copy keeps the buffer, so it must not be released here
IF NOT bInCopyCode AND _pString <> 0 THEN
	__DELETE(_pString);
	_pString := 0;
END_IF
END_METHOD

//FB_Init is always available implicitly and it is used primarily for initialization.
//The return value is not evaluated. For a specific influence, you can also declare the
//methods explicitly and provide additional code there with the standard initialization
//code. You can evaluate the return value.
METHOD FB_Init: BOOL
VAR_INPUT
	bInitRetains: BOOL; // TRUE: the retain variables are initialized (reset warm / reset cold)
	bInCopyCode: BOOL;  // TRUE: the instance will be copied to the copy code afterward (online change)
	url: T_MaxString;  // full endpoint URL, e.g. 'http://192.168.1.10:4318/v1/logs'
	bNoServerCertCheck: BOOL := FALSE;  // allow HTTPS connections to servers with self-signed certificates
END_VAR
THIS^.currentState := E_HttpExporterState.idle;
THIS^._computedState := E_HttpExporterState.idle;

THIS^._urlParsed := F_ParseHttpUrl(url:=url, endpoint=>THIS^._endpoint);

THIS^._client.sHostName := THIS^._endpoint.host;
THIS^._client.nHostPort := THIS^._endpoint.port;
THIS^._client.bKeepAlive := TRUE;
THIS^._client.tConnectionTimeout := T#10S;
IF THIS^._endpoint.useTls THEN
	THIS^._client.stTLS.bNoServerCertCheck := bNoServerCertCheck;
END_IF

THIS^._request.sContentType := 'application/json';
END_METHOD

METHOD isBusy : BOOL
isBusy := THIS^._exportActive;
END_METHOD

METHOD tick : BOOL
VAR_OUTPUT
	failureReason: E_LogRecordExporterFailureReason;
END_VAR
tick := TRUE;
failureReason := E_LogRecordExporterFailureReason.NA;

_execute := THIS^._exportActive;
_execRTrig(CLK := _execute AND_THEN THIS^._records.count > 0);

CASE currentState OF
	E_HttpExporterState.idle:
		IF _execRTrig.Q THEN
			_failureReason := E_LogRecordExporterFailureReason.NA;
			_serializationFailureReason := E_ProtoJsonSerializerFailureReason.NA;
			IF NOT THIS^._urlParsed THEN
				_failureReason := E_LogRecordExporterFailureReason.HTTP_URL_PARSE_FAILURE;
				_computedState := E_HttpExporterState.error;
			ELSE
				_computedState := E_HttpExporterState.serializing;
			END_IF
		END_IF

	E_HttpExporterState.serializing:
		// Serialize the batch and buffer the LogsData document as a byte array payload.
		IF NOT _serializer.serializeLogsData(
			logRecords:=THIS^._records,
			failureReason=>_serializationFailureReason
		) THEN
			_failureReason := E_LogRecordExporterFailureReason.SERIALIZATION_FAILURE;
			_computedState := E_HttpExporterState.error;
		ELSE
			_jsonVal := _serializer.jsonValue;
			IF _jsonVal = 0 OR_ELSE NOT _serializer.parser.IsObject(_jsonVal) THEN
				_failureReason := E_LogRecordExporterFailureReason.SERIALIZATION_FAILURE;
				_computedState := E_HttpExporterState.error;
			ELSE
				_len := _serializer.parser.GetJsonLength(_jsonVal);  // includes the null terminating character
				IF _len = 0 THEN
					_failureReason := E_LogRecordExporterFailureReason.SERIALIZATION_FAILURE;
					_computedState := E_HttpExporterState.error;
				ELSE
					_pString := __NEW(BYTE, _len);
					IF _pString = 0 THEN
						_failureReason := E_LogRecordExporterFailureReason.BUFFER_ALLOCATION_FAILURE;
						_computedState := E_HttpExporterState.error;
					ELSE
						_serializer.parser.CopyJson(_jsonVal, _pString^, _len);
						_computedState := E_HttpExporterState.sending;
					END_IF
				END_IF
			END_IF
		END_IF

	E_HttpExporterState.sending:
		IF NOT _request.bBusy THEN
			IF _request.SendRequest(
				sUri := THIS^._endpoint.path,
				fbClient := THIS^._client,
				eRequestType := ETcIotHttpRequestType.HTTP_POST,
				pContent := _pString,
				nContentSize := _len - 1,
				fbHeader := THIS^._header
			) THEN
				_computedState := E_HttpExporterState.waiting;
			ELSE
				IF _pString <> 0 THEN __DELETE(_pString); _pString := 0; END_IF
				_failureReason := E_LogRecordExporterFailureReason.HTTP_REQUEST_FAILURE;
				_computedState := E_HttpExporterState.error;
			END_IF
		END_IF

	E_HttpExporterState.waiting:
		IF NOT _request.bBusy THEN
			_computedState := E_HttpExporterState.processing;
		END_IF

	E_HttpExporterState.processing:
		IF _request.bError THEN
			IF _pString <> 0 THEN __DELETE(_pString); _pString := 0; END_IF
			_failureReason := E_LogRecordExporterFailureReason.HTTP_REQUEST_FAILURE;
			_computedState := E_HttpExporterState.error;
		ELSE
			statusCode := _request.nStatusCode;
			IF statusCode < 200 OR_ELSE statusCode >= 300 THEN
				IF _pString <> 0 THEN __DELETE(_pString); _pString := 0; END_IF
				_failureReason := E_LogRecordExporterFailureReason.HTTP_STATUS_FAILURE;
				_computedState := E_HttpExporterState.error;
			ELSE
				IF _pString <> 0 THEN __DELETE(_pString); _pString := 0; END_IF
				_computedState := E_HttpExporterState.done;
			END_IF
		END_IF

	E_HttpExporterState.done:
		IF NOT _execute THEN
			_computedState := E_HttpExporterState.idle;
		END_IF
		THIS^.free();

	E_HttpExporterState.error:
		// Retain the failure until export accepts a new batch.
END_CASE

currentState := _computedState;

IF currentState = E_HttpExporterState.done
	OR_ELSE currentState = E_HttpExporterState.error THEN
	THIS^.free();
END_IF

THIS^._client.Execute();

IF currentState = E_HttpExporterState.error THEN
	tick := FALSE;
	failureReason := _failureReason;
END_IF
END_METHOD

END_FUNCTION_BLOCK

// ---- OTEL/EXPORTING/FUNCTIONS/F_ParseHttpUrl.TcPOU
(*
	Splits a full endpoint URL into scheme, host, port and path, for example
	'http://192.168.1.10:4318/v1/traces'. The scheme must be lower-case http or https, and
	IPv6 hosts are not supported. Returns FALSE when the URL cannot be parsed; endpoint then
	holds no usable host.
*)
FUNCTION F_ParseHttpUrl : BOOL
VAR_INPUT
	url: T_MaxString;
END_VAR
VAR_OUTPUT
	endpoint: ST_HttpEndpoint;
END_VAR
VAR
	_rest: T_MaxString;
	_portString: T_MaxString;
	_pathStart: INT;
	_colonIdx: INT;
END_VAR

F_ParseHttpUrl := FALSE;
endpoint.useTls := FALSE;
endpoint.host := '';
endpoint.port := 0;
endpoint.path := '/';

IF FIND(url, 'https://') = 1 THEN
	endpoint.useTls := TRUE;
	_rest := RIGHT(url, LEN(url) - 8);
ELSIF FIND(url, 'http://') = 1 THEN
	endpoint.useTls := FALSE;
	_rest := RIGHT(url, LEN(url) - 7);
ELSE
	RETURN;
END_IF

_pathStart := FIND(_rest, '/');
IF _pathStart > 0 THEN
	endpoint.host := LEFT(_rest, _pathStart - 1);
	endpoint.path := RIGHT(_rest, LEN(_rest) - _pathStart + 1);
ELSE
	endpoint.host := _rest;
	endpoint.path := '/';
END_IF

IF endpoint.useTls THEN
	endpoint.port := 443;
ELSE
	endpoint.port := 80;
END_IF

_colonIdx := FIND(endpoint.host, ':');
IF _colonIdx > 0 THEN
	_portString := RIGHT(endpoint.host, LEN(endpoint.host) - _colonIdx);
	IF _portString = '' THEN RETURN; END_IF
	endpoint.port := STRING_TO_UINT(_portString);
	IF endpoint.port = 0 THEN RETURN; END_IF
	endpoint.host := LEFT(endpoint.host, _colonIdx - 1);
END_IF

IF endpoint.host = '' THEN RETURN; END_IF

F_ParseHttpUrl := TRUE;

END_FUNCTION

// ---- OTEL/LOGGING/LOGGER/FUNCTION_BLOCKS/FB_Logger.TcPOU
{attribute 'enable_dynamic_creation'}
FUNCTION_BLOCK FB_Logger
VAR_OUTPUT
	pLogRecord: POINTER TO FB_LogRecord;
END_VAR
VAR
	_scope: REFERENCE TO FB_InstrumentationScope;
	_provider: REFERENCE TO FB_LoggerProvider;
	_failed: BOOL;
	_failureReason: E_LoggerFailureReason;
END_VAR

METHOD _createLogRecord : BOOL
VAR_IN_OUT
	pDest: POINTER TO FB_LogRecord;
END_VAR
VAR_INPUT
	severityNumber: E_SeverityNumber;
	timestamp: ULINT;
END_VAR
VAR_OUTPUT
	failureReason: E_LoggerFailureReason;
END_VAR
VAR
	_logRecord: POINTER TO FB_LogRecord;
	_attributesFailureResult: E_AttributesFailureReason;
END_VAR
_createLogRecord := FALSE;
failureReason := E_LoggerFailureReason.NA;

IF pDest <> 0 THEN
	failureReason := E_LoggerFailureReason.LOG_RECORD_ALREADY_STARTED;
	RETURN;
END_IF

_logRecord := __NEW(FB_LogRecord(
	severityNumber:=severityNumber,
	timestamp:=timestamp
));

IF _logRecord = 0 THEN
	failureReason := E_LoggerFailureReason.MEMORY_ALLOCATION_FAILURE;
	RETURN;
END_IF

IF NOT _logRecord^.resource.copyFrom(src:=THIS^.resource, failureResult=>_attributesFailureResult) THEN
	IF _attributesFailureResult = E_AttributesFailureReason.MEMORY_ALLOCATION_FAILURE THEN
		failureReason := E_LoggerFailureReason.MEMORY_ALLOCATION_FAILURE;
	ELSE
		failureReason := E_LoggerFailureReason.SNAPSHOT_COPY_FAILURE;
	END_IF
	_logRecord^.delete(pSelf:=_logRecord);
	RETURN;
END_IF

IF NOT _logRecord^.scope.copyFrom(src:=THIS^.scope, failureResult=>_attributesFailureResult) THEN
	IF _attributesFailureResult = E_AttributesFailureReason.MEMORY_ALLOCATION_FAILURE THEN
		failureReason := E_LoggerFailureReason.MEMORY_ALLOCATION_FAILURE;
	ELSE
		failureReason := E_LoggerFailureReason.SNAPSHOT_COPY_FAILURE;
	END_IF
	_logRecord^.delete(pSelf:=_logRecord);
	RETURN;
END_IF

pDest := _logRecord;
_logRecord := 0;
_createLogRecord := failureReason = E_LoggerFailureReason.NA;
END_METHOD

METHOD _shouldReturnEarly : BOOL
_shouldReturnEarly := TRUE;

// Preserve the first failure in the active fluent chain.
IF THIS^._failed THEN
	RETURN;
END_IF

// fail early if the log record hasn't been built
IF THIS^.pLogRecord = 0 THEN
	THIS^._failed := TRUE;
	THIS^._failureReason := E_LoggerFailureReason.LOG_RECORD_NOT_STARTED;
	RETURN;
END_IF

_shouldReturnEarly := FALSE;
END_METHOD

(*
	Function emits a log record by pushing it to the owning provider's queue.
	Each log record owns a snapshot of its instrumentation scope and resource, so processors
	may retain the record after its logger or provider has been destroyed.
*)
METHOD emit: BOOL
VAR_OUTPUT
	failureResult: E_LoggerFailureReason;
END_VAR
emit := FALSE;
failureResult := E_LoggerFailureReason.NA;

// Preserve the first fluent method failure while releasing the incomplete record.
IF THIS^._failed THEN
	IF THIS^.pLogRecord <> 0 THEN THIS^.pLogRecord^.delete(pSelf:=THIS^.pLogRecord); END_IF
	failureResult := THIS^._failureReason;
	RETURN;
END_IF

IF THIS^.pLogRecord = 0 THEN
	THIS^._failed := TRUE;
	THIS^._failureReason := E_LoggerFailureReason.LOG_RECORD_NOT_STARTED;
	failureResult := THIS^._failureReason;
	RETURN;
END_IF

// Push the record to the provider's queue for cyclical processing.
IF NOT THIS^._provider.onEmit(THIS^.pLogRecord) THEN
	THIS^.pLogRecord^.delete(pSelf:=THIS^.pLogRecord);
	THIS^._failed := TRUE;
	THIS^._failureReason := E_LoggerFailureReason.TRANSFER_TO_PROVIDER_FAILURE;
	failureResult := THIS^._failureReason;
	RETURN;
END_IF

emit := THIS^._failureReason = E_LoggerFailureReason.NA;
THIS^._failed := FALSE;
THIS^._failureReason := E_LoggerFailureReason.NA;
END_METHOD

//FB_Exit must be implemented explicitly. If there is an implementation, then the
//method is called before the controller removes the code of the function block instance
//(implicit call). The return value is not evaluated.
METHOD FB_Exit: BOOL
VAR_INPUT
    bInCopyCode: BOOL;  // TRUE: the exit method is called in order to leave the instance which will be copied afterwards (online change).
END_VAR
// during an online change the copied instance keeps pLogRecord, so the record must survive
IF NOT bInCopyCode THEN
	THIS^.free();
END_IF
END_METHOD

//FB_Init is always available implicitly and it is used primarily for initialization.
//The return value is not evaluated. For a specific influence, you can also declare the
//methods explicitly and provide additional code there with the standard initialization
//code. You can evaluate the return value.
METHOD FB_Init: BOOL
VAR_INPUT
    bInitRetains: BOOL; // TRUE: the retain variables are initialized (reset warm / reset cold)
    bInCopyCode: BOOL;  // TRUE: the instance will be copied to the copy code afterward (online change)
	scope: REFERENCE TO FB_InstrumentationScope;
	provider: REFERENCE TO FB_LoggerProvider;
END_VAR
THIS^._scope REF= scope;
THIS^._provider REF= provider;
END_METHOD

METHOD free
VAR_INPUT
END_VAR
IF THIS^.pLogRecord <> 0 THEN
	THIS^.pLogRecord^.delete(pSelf:=THIS^.pLogRecord);
END_IF
THIS^._failed := TRUE;
THIS^._failureReason := E_LoggerFailureReason.LOG_RECORD_NOT_STARTED;
END_METHOD

METHOD reset
VAR_INPUT
END_VAR
THIS^.free();
THIS^._failed := FALSE;
THIS^._failureReason := E_LoggerFailureReason.NA;
END_METHOD

PROPERTY resource : REFERENCE TO FB_Resource
GET
resource REF= THIS^._provider.resource;
END_GET
END_PROPERTY

PROPERTY scope : REFERENCE TO FB_InstrumentationScope
GET
scope REF= THIS^._scope;
END_GET
END_PROPERTY

METHOD setBody: REFERENCE TO FB_Logger
VAR_INPUT
	str: T_MaxString;  // use setBody_AnyValue if the body isn't a string
END_VAR
VAR
	_pDest: POINTER TO FB_String;
	_factoryFailureReason: E_ValueFactoryFailureReason;
END_VAR
setBody REF= THIS^;

IF THIS^._shouldReturnEarly() THEN
	RETURN;
END_IF

// Create an owned string body.
IF NOT ValueFactory.createString(
	pDest:=_pDest,
	pString:=ADR(str),
	failureReason=>_factoryFailureReason
	) THEN
	THIS^._failed := TRUE;
	IF _factoryFailureReason = E_ValueFactoryFailureReason.MEMORY_ALLOCATION_FAILURE THEN
		THIS^._failureReason := E_LoggerFailureReason.MEMORY_ALLOCATION_FAILURE;
	ELSE
		THIS^._failureReason := E_LoggerFailureReason.BODY_VALUE_INVALID;
	END_IF
	RETURN;
END_IF

// Replace the body only after the new value has been created successfully.
IF THIS^.pLogRecord^.body <> 0 THEN
	THIS^.pLogRecord^.body^.delete(pSelf:=THIS^.pLogRecord^.body);
END_IF
THIS^.pLogRecord^.body := _pDest;
_pDest := 0;
END_METHOD

METHOD setBody_AnyValue: REFERENCE TO FB_Logger
VAR_INPUT
	pVal: POINTER TO FB_AnyValue;  // use setBody_AnyValue if the body isn't a string
END_VAR
VAR
	_pDest: POINTER TO FB_AnyValue;
	_factoryFailureReason: E_ValueFactoryFailureReason;
END_VAR
setBody_AnyValue REF= THIS^;

IF THIS^._shouldReturnEarly() THEN
	RETURN;
END_IF

// check that the value is valid
IF pVal = 0 THEN
	THIS^._failed := TRUE;
	THIS^._failureReason := E_LoggerFailureReason.BODY_VALUE_POINTER_NULL;
	RETURN;
END_IF

// try to create a clone
IF NOT ValueFactory.cloneAnyValue(
	pDest:=_pDest,
	pSrc:=pVal,
	failureReason=>_factoryFailureReason
	) THEN
	THIS^._failed := TRUE;
	CASE _factoryFailureReason OF
		E_ValueFactoryFailureReason.MEMORY_ALLOCATION_FAILURE:
			THIS^._failureReason := E_LoggerFailureReason.MEMORY_ALLOCATION_FAILURE;
		E_ValueFactoryFailureReason.UNSUPPORTED_VALUE_TYPE:
			THIS^._failureReason := E_LoggerFailureReason.BODY_VALUE_TYPE_UNSUPPORTED;
	ELSE
		THIS^._failureReason := E_LoggerFailureReason.BODY_VALUE_INVALID;
	END_CASE
	RETURN;
END_IF

// clean up the prior record if it existed
IF THIS^.pLogRecord^.body <> 0 THEN
	THIS^.pLogRecord^.body^.delete(pSelf:=THIS^.pLogRecord^.body);
END_IF
// transfer ownership
THIS^.pLogRecord^.body := _pDest;
_pDest := 0;
END_METHOD

METHOD setEventName: REFERENCE TO FB_Logger
VAR_INPUT
	str: T_MaxString;
END_VAR
VAR
	_pDest: POINTER TO FB_String;
	_factoryFailureReason: E_ValueFactoryFailureReason;
END_VAR
setEventName REF= THIS^;

IF THIS^._shouldReturnEarly() THEN
	RETURN;
END_IF

// create FB_String
IF NOT ValueFactory.createString(
	pDest:=_pDest,
	pString:=ADR(str),
	failureReason=>_factoryFailureReason
	) THEN
	THIS^._failed := TRUE;
	IF _factoryFailureReason = E_ValueFactoryFailureReason.MEMORY_ALLOCATION_FAILURE THEN
		THIS^._failureReason := E_LoggerFailureReason.MEMORY_ALLOCATION_FAILURE;
	ELSE
		THIS^._failureReason := E_LoggerFailureReason.EVENT_NAME_INVALID;
	END_IF
	RETURN;
END_IF

// assign to record event name
// delete old event name if it exists
IF THIS^.pLogRecord^.eventName <> 0 THEN
	THIS^.pLogRecord^.eventName^.delete(pSelf:=THIS^.pLogRecord^.eventName);
END_IF
// transfer ownership of the pointer
THIS^.pLogRecord^.eventName := _pDest;
_pDest := 0;
END_METHOD

(*
	Fills the record's trace context from the span: the trace id, span id and W3C trace flags, the parts of the
	span context that the log data model carries. Trace state and remoteness are not copied.
	The log then correlates with the span and carries its sampled bit. The span is borrowed for the call only.
	A null span, or a span without ids, is a no-op rather than a failure, so the same chain works inside and outside a span.
*)
METHOD setTraceContextFromSpan: REFERENCE TO FB_Logger
VAR_INPUT
	pSpan: POINTER TO FB_Span;
END_VAR
setTraceContextFromSpan REF= THIS^;

IF THIS^._shouldReturnEarly() THEN
	RETURN;
END_IF

// every span has both ids, so a span without them is not worth failing the log over
IF pSpan = 0 OR_ELSE pSpan^.traceId = 0 OR_ELSE pSpan^.spanId = 0 THEN
	RETURN;
END_IF

THIS^._setTraceId(pBytes:=ADR(pSpan^.traceId^.bytes), nSize:=SIZEOF(pSpan^.traceId^.bytes));
THIS^._setSpanId(pBytes:=ADR(pSpan^.spanId^.bytes), nSize:=SIZEOF(pSpan^.spanId^.bytes));
// bits 0-7 of the span flags are the W3C trace flags, the rest describe the parent and stay on the span
THIS^._setFlags(traceFlags:=TO_BYTE(pSpan^.flags AND TO_UDINT(E_SpanFlags.SPAN_FLAGS_TRACE_FLAGS_MASK)));
END_METHOD

METHOD setNumberAttribute: REFERENCE TO FB_Logger
VAR_INPUT
	key: T_MaxString;
	value: ANY_NUM;
END_VAR
VAR
	_attributesSuccess: BOOL;
	_attributesFailureReason: E_AttributesFailureReason;
END_VAR
setNumberAttribute REF= THIS^;

IF THIS^._shouldReturnEarly() THEN
	RETURN;
END_IF

_attributesSuccess := THIS^.pLogRecord^.attributes.setNumberAttribute_AnyType(
	key:=key,
	value:=value,
	failureReason=>_attributesFailureReason
);
IF NOT _attributesSuccess THEN
	THIS^._failed := TRUE;
	CASE _attributesFailureReason OF
		E_AttributesFailureReason.MEMORY_ALLOCATION_FAILURE:
			THIS^._failureReason := E_LoggerFailureReason.MEMORY_ALLOCATION_FAILURE;
		E_AttributesFailureReason.ATTRIBUTE_COUNT_LIMIT_REACHED:
			THIS^._failureReason := E_LoggerFailureReason.ATTRIBUTE_COUNT_LIMIT_REACHED;
		E_AttributesFailureReason.KV_VALUE_TYPE_UNSUPPORTED:
			THIS^._failureReason := E_LoggerFailureReason.ATTRIBUTE_VALUE_TYPE_UNSUPPORTED;
	ELSE
		THIS^._failureReason := E_LoggerFailureReason.ATTRIBUTE_VALUE_INVALID;
	END_CASE
END_IF
END_METHOD

(*
	Sets the record's W3C trace flags; bit 0 is sampled. Application code uses setTraceContextFromSpan; this setter is
	for tests and for setTraceContextFromSpan itself. A BYTE keeps the reserved bits 8-31 of the record's flags zero.
*)
METHOD _setFlags: REFERENCE TO FB_Logger
VAR_INPUT
	traceFlags: BYTE;
END_VAR
_setFlags REF= THIS^;

IF THIS^._shouldReturnEarly() THEN
	RETURN;
END_IF

THIS^.pLogRecord^.flags := TO_UDINT(traceFlags);
END_METHOD

(* Sets the record's span id from raw bytes. Application code uses setTraceContextFromSpan; this setter is for tests and for setTraceContextFromSpan itself. *)
METHOD _setSpanId: REFERENCE TO FB_Logger
VAR_INPUT
	pBytes: POINTER TO BYTE;
	nSize: UDINT;
END_VAR
VAR
	_pDest: POINTER TO FB_SpanId;
	_factoryFailureReason: E_ValueFactoryFailureReason;
END_VAR
_setSpanId REF= THIS^;

IF THIS^._shouldReturnEarly() THEN
	RETURN;
END_IF

// create an instance of FB_SpanId
IF NOT ValueFactory.createSpanId(
	pDest:=_pDest,
	pBytes:=pBytes,
	nSize:=nSize,
	failureReason=>_factoryFailureReason
	) THEN
	THIS^._failed := TRUE;
	CASE _factoryFailureReason OF
		E_ValueFactoryFailureReason.MEMORY_ALLOCATION_FAILURE:
			THIS^._failureReason := E_LoggerFailureReason.MEMORY_ALLOCATION_FAILURE;
		E_ValueFactoryFailureReason.SPAN_ID_BYTES_POINTER_NULL:
			THIS^._failureReason := E_LoggerFailureReason.SPAN_ID_BYTES_POINTER_NULL;
		E_ValueFactoryFailureReason.SPAN_ID_BYTE_COUNT_TOO_SMALL:
			THIS^._failureReason := E_LoggerFailureReason.SPAN_ID_BYTE_COUNT_TOO_SMALL;
	ELSE
		THIS^._failureReason := E_LoggerFailureReason.SPAN_ID_INVALID;
	END_CASE
	RETURN;
END_IF

// assign to the record
// delete the prior record if it exists
IF THIS^.pLogRecord^.spanId <> 0 THEN
	THIS^.pLogRecord^.spanId^.delete(pSelf:=THIS^.pLogRecord^.spanId);
END_IF
// transfer owneship of the data
THIS^.pLogRecord^.spanId := _pDest;
_pDest := 0;
END_METHOD

METHOD setStringAttribute: REFERENCE TO FB_Logger
VAR_INPUT
	key: T_MaxString;
	value: T_MaxString;
END_VAR
VAR
	_attributesSuccess: BOOL;
	_attributesFailureReason: E_AttributesFailureReason;
END_VAR
setStringAttribute REF= THIS^;

IF THIS^._shouldReturnEarly() THEN
	RETURN;
END_IF

